RoboDK station: 2026-11-5.rdk

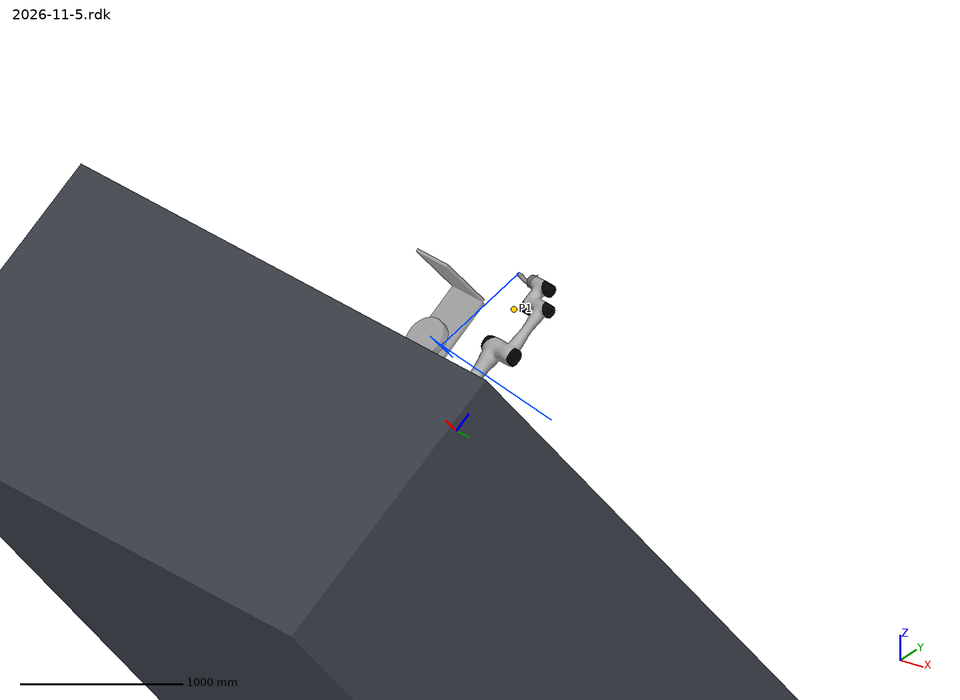
[picture v0: the station drawn from its stored meshes, robots at their saved joint values, targets as dots, program paths as lines]
Station 新建工作站 (1) (saved by RoboDK 5.9.0). Poses are relative to the parent item; angles as X-Y-Z fixed-axis rotations.
Station parameters (name, value as stored): Trace_Render_Style, 0
  - Python program TCP真实运动_升级前备份_20260910_170410 (listed below)
  - Python program 方向角计算 (listed below)
  - Python program test (listed below)
  - Python program 机械臂法兰真实运动_改名修复前_20261014_114144_改名修复前_20261014_114144 (listed below)
  - Python program TCP真实运动_到位复核前备份_20260910_172919 (listed below)
  - Python program TCP真实运动_改名修复前_20261014_114144 (listed below)
  - program _probe_P11 (4 instructions, listed below)
  - Python program 机械臂法兰真实运动 (listed below)
  - Python program TCP仿真 (listed below)
  - Python program TCP真实运动_偏离50版_20261009_142831 (listed below)
  - Python program TCP真实运动_偏离50版_20261009_144043 (listed below)
  - Python program TCP真实运动 (listed below)
  - Python program TCP真实运动_P2P版_修复前_v14w40_20261027 (listed below)
  - Python program TCP真实运动_P2P版_优化前_v14w41_20261027 (listed below)
  - frame Dobot CR5 Base_控制器对齐 at (346.03, 1005.01, 515.52) mm, rotated rx 1.05 ry -48.85 rz -107.35 deg
    - robot Dobot CR5: 6 axes, payload 5 kg, reach 900 mm, repeatability 0.03 mm, weight 23 kg
        modified DH rows (alpha deg, a mm, theta deg, d mm): 0, 0, 0, 147; 90.028, 0.839, 90, 0; -0.44, 427.688, 0, 0; 0.304, 357.005, -90, 140.421; -90.09, 0.126, 0, 115.885; 89.829, 0.736, 180, 104.5
        joint limits [-360, -360, -160, -360, -360, -360] to [360, 360, 160, 360, 360, 360]; home [0, 0, -90, 90, 90, 0]; saved at [0, 0, 0, 0, 0, 0]
      - tool CR5_TCP_126mm, TCP at (0, 0, 126) mm
      - tool _CR5_FLANGE_DIRECT_TEMP, TCP at (0, 0, 0) mm
      - tool _, TCP at (0, 0, 130) mm
      - tool CR5_TCP_130mm, TCP at (0, 0, 130) mm
      - tool _offline_TCP130_test, TCP at (0, 0, 130) mm
      - object  at (0, 0, 0) mm, size 120.1 x 130 x 24.6 mm, geometry from handle130.stl
    - target P1 (joint target) at (-20.1, -241.48, 846.75) mm, rotated rx -90 ry 1.35 rz 179.96 deg; joints [0, -37.451, 84.112, -46.661, 0, 0] of Dobot CR5
    - object  at (0, 0, 0) mm, rotated rx 0 ry -1.35 rz -0.05 deg, size 650 x 650 x 80 mm
    - object  at (0, 0, 0) mm, rotated rx 0 ry -1.35 rz -0.05 deg, size 4000 x 4000 x 2000 mm
    - object  at (0, 223.9, 120) mm, size 450 x 300 x 750 mm, geometry from baffle_semiopen_3face_y300.stl
    - object  at (0, -692.1, 420) mm, rotated rx 90 ry 0 rz 90 deg, size 280 x 280 x 50 mm, geometry from cylinder_R140_H50.stl
  - Python program TCP真实运动_P2P版_16稳定版_替换前_20261104_095940 (listed below)
  - program _TCP仿真_路径预检 (0 instructions, listed below)
  - Python program TCP真实运动_P2P版 (listed below)
  - program 轨迹17_仿真27点 (30 instructions, listed below)
  - object  at (0, 0, 0) mm
  - Python program CR5_零位到P1_上传 (listed below)
  - Python program CR5_首段MoveL_上传 (listed below)
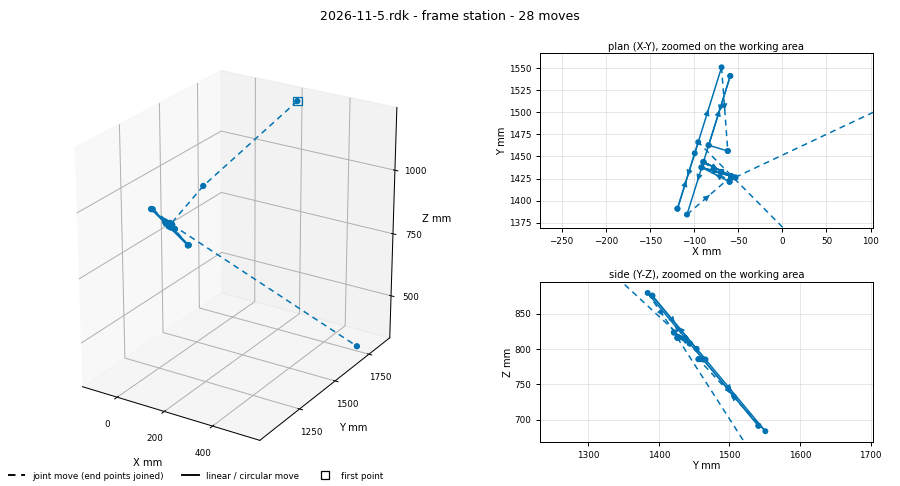
[picture p0: tool path of 2026-11-5.rdk in frame station, 28 of 30 moves have a stored position in this frame; points joined in program order, loops and branches not executed]

--- Python program TCP真实运动_升级前备份_20260910_170410 ---
# -*- coding: utf-8 -*-
"""
RoboDK 实机运动控制（基于 robodk_movej_diag.py 的成功模式）
- 单点：TCP 输入 -> IK 检测 -> MoveL/MoveJ 执行
- 连续轨迹：坐标列表 -> 逐点 IK 检测 -> MoveJ+MoveL 序列
模式：RUNMODE_RUN_ROBOT + robot.Connect()
"""

from robodk.robolink import *
from robodk.robomath import *
import tkinter as tk
from tkinter import ttk, scrolledtext, filedialog
import time
import math
import json

ROBOT_SPEED = 20.0
NL = chr(10)

RDK = Robolink()

def fanuc_to_pose(x, y, z, rx, ry, rz):
    return Fanuc_2_Pose([x, y, z, rx, ry, rz])

def pose_to_fanuc(pose):
    return Pose_2_Fanuc(pose)

# ---- 获取机器人 ----
robot = RDK.Item('', ITEM_TYPE_ROBOT)
if not robot.Valid():
    raise Exception("未找到机器人")

# ---- 全局变量 ----
text_points = None
text_log = None
record_text = None
entries_single = None
entries_joint = None
move_type = None
trajectory_records = []
_connected = False

# ============================================================
# 日志
# ============================================================
def log(s):
    print(s)
    if text_log:
        text_log.insert(tk.END, str(s) + NL)
        text_log.see(tk.END)
        root.update_idletasks()

# ============================================================
# 连接（只连一次，复用）
# ============================================================
def ensure_connected():
    global _connected
    if _connected:
        return True
    try:
        robot.Connect()
        time.sleep(1.5)
        status, msg = robot.ConnectedState()
        log("连接状态: %s, %s" % (status, msg))
        RDK.setRunMode(RUNMODE_RUN_ROBOT)
        log("RunMode: %s" % RDK.RunMode())
        if status < 0:
            _connected = False
            log("机器人连接未建立，状态=%s：%s" % (status, msg))
            return False
        _connected = True
        return True
    except Exception as e:
        log("连接失败: %s" % e)
        return False

# ============================================================
# 解析坐标
# ============================================================
def parse_points():
    if not text_points:
        return []
    raw = text_points.get("1.0", tk.END)
    points = []
    for line in raw.strip().split(NL):
        line = line.strip()
        if not line or line.startswith("#"):
            continue
        try:
            vals = [float(v.strip()) for v in line.split(",")]
            if len(vals) >= 6:
                points.append(vals[:6])
        except ValueError:
            pass
    return points

# ============================================================
# 读取当前位置
# ============================================================
def read_current(entries=None):
    try:
        pose = robot.Pose()
        v = pose_to_fanuc(pose)
        log("")
        log("当前 TCP：X=%.3f Y=%.3f Z=%.3f Rx=%.3f Ry=%.3f Rz=%.3f" % tuple(v[:6]))
    except Exception as e:
        log("读取失败：%s" % e)

def fill_current(entries=None):
    try:
        pose = robot.Pose()
        v = pose_to_fanuc(pose)
        if entries:
            for e, val in zip(entries, v):
                e.delete(0, tk.END)
                e.insert(0, "%.3f" % val)
        log("当前 TCP 已填入")
    except Exception as e:
        log("读取失败：%s" % e)

# ============================================================
# IK 检测
# 注意：SolveIK 显式使用当前 Tool + Reference，和 MoveL/MoveJ 保持一致。
# ============================================================
def check_ik_single(entries=None):
    if not entries:
        return
    try:
        values = [float(e.get()) for e in entries]
    except ValueError:
        log("输入无效")
        return

    x, y, z, rx, ry, rz = values
    target = fanuc_to_pose(x, y, z, rx, ry, rz)
    log("")
    log("目标：X=%.3f Y=%.3f Z=%.3f Rx=%.3f Ry=%.3f Rz=%.3f" % (x, y, z, rx, ry, rz))

    try:
        tool_pose = robot.PoseTool()
        frame_pose = robot.PoseFrame()
        joints = robot.SolveIK(target, tool=tool_pose, reference=frame_pose)
        if joints is None:
            log("IK 不可达")
        else:
            q = joints.list()
            if len(q) < 6:
                log("IK 返回关节数量异常：%d，原始数据=%r" % (len(q), q))
                return
            log("IK 可达")
            log("  关节：J1=%.2f J2=%.2f J3=%.2f J4=%.2f J5=%.2f J6=%.2f" % tuple(q[:6]))
    except Exception as e:
        log("检测失败：%s" % e)

def check_all_ik():
    points = parse_points()
    if not points:
        log("没有有效点")
        return

    log("")
    log("========== 检测全部 %d 个点 ==========" % len(points))
    all_ok = True
    for i, p in enumerate(points):
        try:
            target = fanuc_to_pose(*p)
            joints = robot.SolveIK(target, tool=robot.PoseTool(), reference=robot.PoseFrame())
            if joints is None:
                log("  P%d: 不可达" % (i+1))
                all_ok = False
            else:
                q = joints.list()
                if len(q) < 6:
                    raise ValueError("IK 返回关节数量异常: %d, raw=%r" % (len(q), q))
                log("  P%d: 可达  J1=%.1f J2=%.1f J3=%.1f J4=%.1f J5=%.1f J6=%.1f" % (i+1, *q[:6]))
        except Exception as e:
            log("  P%d: 检测失败 %s" % (i+1, e))
            all_ok = False
    if all_ok:
        log("全部 %d 个点可达" % len(points))
    else:
        log("存在不可达点，执行时会跳过")

# ============================================================
# 执行单点
# ============================================================
def execute_single(entries=None, mtype="MoveL"):
    if not entries:
        return
    try:
        values = [float(e.get()) for e in entries]
    except ValueError:
        log("输入无效")
        return

    x, y, z, rx, ry, rz = values
    target = fanuc_to_pose(x, y, z, rx, ry, rz)
    log("")
    log("目标：X=%.3f Y=%.3f Z=%.3f Rx=%.3f Ry=%.3f Rz=%.3f" % (x, y, z, rx, ry, rz))

    try:
        tool_pose = robot.PoseTool()
        frame_pose = robot.PoseFrame()
        joints = robot.SolveIK(target, tool=tool_pose, reference=frame_pose)
        if joints is None:
            log("IK 不可达，取消执行")
            return
        q = joints.list()
        if len(q) < 6:
            log("IK 返回关节数量异常：%d，取消执行；原始数据=%r" % (len(q), q))
            return
        log("IK 可达：J1=%.2f J2=%.2f J3=%.2f J4=%.2f J5=%.2f J6=%.2f" % tuple(q[:6]))
    except Exception as e:
        log("IK 检查失败：%s" % e)
        return

    if not ensure_connected():
        return

    try:
        robot.setPoseFrame(robot.PoseFrame())
        robot.setPoseTool(robot.PoseTool())
        robot.setSpeed(ROBOT_SPEED)
        log("发送 %s..." % mtype)
        if mtype == "MoveJ":
            robot.MoveJ(target)
        else:
            robot.MoveL(target)
        log("执行完成")
    except Exception as e:
        log("失败: %s: %s" % (type(e).__name__, e))

# ============================================================
# 连续运动：选项卡3直接输入 TCP / 关节点，逐点检查后加入轨迹
# ============================================================
trajectory_records = []
record_text = None
traj_entries = None
traj_type = None
singular_var = None
j6_direction_var = None


def _parse_six_from_entries(entries, label):
    if not entries or len(entries) != 6:
        log("%s输入框异常：需要 6 个值" % label)
        return None
    try:
        vals = [float(e.get().strip()) for e in entries]
    except (ValueError, AttributeError):
        log("%s输入无效：6 个值必须全部为数字" % label)
        return None
    if not all(math.isfinite(v) for v in vals):
        log("%s输入无效：不能包含 NaN 或无穷值" % label)
        return None
    return vals


def _check_tcp_reachable(vals):
    """检查单个 TCP 点 IK 是否可达，返回 (True, target, joints)。"""
    try:
        target = fanuc_to_pose(*vals)
        tool_pose = robot.PoseTool()
        frame_pose = robot.PoseFrame()
        joints = robot.SolveIK(target, tool=tool_pose, reference=frame_pose)

        if joints is None:
            log("TCP IK：不可达")
            return False, None, None

        q = joints.list()
        if len(q) < 6:
            log("TCP IK：返回关节数量异常：%r" % q)
            return False, None, None

        log("TCP IK：可达")
        log("  IK关节：J1=%.2f J2=%.2f J3=%.2f J4=%.2f J5=%.2f J6=%.2f" % tuple(q[:6]))
        return True, target, q[:6]
    except Exception as e:
        log("TCP IK 检查失败：%s: %s" % (type(e).__name__, e))
        return False, None, None


def _check_tcp_segment_continuous(prev_vals, curr_vals, segment_index, samples=20):
    """检查前一个 TCP 点到当前 TCP 点之间的整段插补路径 IK 连续可达性。

    暂不考虑障碍物，只对 TCP 位姿做线性插值，并对每个采样位姿执行 SolveIK。
    起点和终点也包含在采样检查中。
    """
    if prev_vals is None:
        return True

    log("开始检查 P%d -> P%d 的 TCP 连续 IK（%d 个采样点）" %
        (segment_index - 1, segment_index, samples + 1))

    tool_pose = robot.PoseTool()
    frame_pose = robot.PoseFrame()

    for k in range(samples + 1):
        t = float(k) / float(samples)
        vals = [prev_vals[i] + (curr_vals[i] - prev_vals[i]) * t for i in range(6)]
        try:
            pose = fanuc_to_pose(*vals)
            joints = robot.SolveIK(pose, tool=tool_pose, reference=frame_pose)
            if joints is None:
                log("  P%d -> P%d：第 %d/%d 个采样点 IK 不可达，t=%.3f" %
                    (segment_index - 1, segment_index, k + 1, samples + 1, t))
                log("  TCP：X=%.3f Y=%.3f Z=%.3f Rx=%.3f Ry=%.3f Rz=%.3f" % tuple(vals))
                return False
            q = joints.list()
            if len(q) < 6:
                log("  P%d -> P%d：第 %d 个采样点 IK 返回异常：%r" %
                    (segment_index - 1, segment_index, k + 1, q))
                return False
        except Exception as e:
            log("  P%d -> P%d：第 %d 个采样点 IK 检查失败：%s: %s" %
                (segment_index - 1, segment_index, k + 1, type(e).__name__, e))
            return False

    log("P%d -> P%d：连续 IK 检查通过" % (segment_index - 1, segment_index))
    return True


def _check_joint_reachable(q):
    """兼容旧代码：关节点不做可达性/限位检查，输入合法即可加入。"""
    return True


def refresh_record_list():
    if record_text is None:
        return

    record_text.delete("1.0", tk.END)

    for i, rec in enumerate(trajectory_records, 1):
        kind = rec["type"]
        vals = rec["values"]

        if kind == "TCP":
            mark = " [J6特异点 %s180°]" % ("+" if rec.get("j6_delta", 180) >= 0 else "-") if rec.get("singular", False) else ""
            record_text.insert(
                tk.END,
                "P%-3d [TCP]%s   X=%9.3f Y=%9.3f Z=%9.3f Rx=%8.3f Ry=%8.3f Rz=%8.3f%s" %
                (i, mark, *vals, NL)
            )
        else:
            record_text.insert(
                tk.END,
                "P%-3d [JNT]   J1=%8.3f J2=%8.3f J3=%8.3f J4=%8.3f J5=%8.3f J6=%8.3f%s" %
                (i, *vals, NL)
            )


def add_and_check_trajectory_point():
    """
    选项卡3逐点输入：
    - 普通 TCP：立即做端点 IK，并检查与前一个普通 TCP 点之间的连续 IK。
    - TCP 末端特异点：跳过 IK；要求与前一个普通 TCP 点 XYZ 相同，执行时仅 J6 转 ±180°。
    - 关节：不做 IK/限位检查，只将角度规范到 (-180°, 180°]。
    注意：这些检查只在“加入点”时完成；正式实机执行时不再做轨迹预检。
    """
    kind = traj_type.get()
    vals = _parse_six_from_entries(traj_entries, kind)
    if vals is None:
        return

    log("")
    log("========== 检查连续运动第 %d 点 ==========" % (len(trajectory_records) + 1))

    is_singular = bool(singular_var.get()) if (kind == "TCP" and singular_var is not None) else False
    j6_delta = int(j6_direction_var.get()) if (j6_direction_var is not None) else 180

    if kind == "TCP" and is_singular:
        if not trajectory_records:
            log("末端特异点不能作为第一个点：需要先有一个起始运动点。")
            return
        prev = trajectory_records[-1]
        if prev["type"] != "TCP" or prev.get("singular", False):
            log("末端特异点前一项必须是普通 TCP 点。")
            return
        prev_vals = prev["values"]
        pos_err = math.sqrt(sum((vals[k] - prev_vals[k]) ** 2 for k in range(3)))
        if pos_err > 1e-3:
            log("末端特异点未加入：XYZ 必须与前一个普通 TCP 点相同。")
            log("  与前一点位置差：%.6f mm" % pos_err)
            return
        try:
            target = fanuc_to_pose(*vals)
        except Exception as e:
            log("末端特异点姿态转换失败：%s: %s" % (type(e).__name__, e))
            return

        trajectory_records.append({
            "type": "TCP", "values": vals[:], "target": target, "joints": None,
            "singular": True, "j6_delta": j6_delta,
        })
        log("P%d [TCP-特异点]：已加入，跳过 IK。" % len(trajectory_records))
        log("  执行时保持 J1~J5 不变，仅让 J6 转 %+d°。" % j6_delta)
        if singular_var is not None:
            singular_var.set(False)
        refresh_record_list()
        return

    if kind == "TCP":
        ok, target, joints = _check_tcp_reachable(vals)
        if not ok:
            log("该 TCP 点未加入轨迹。")
            return

        # 只在点加入阶段检查连续 IK；实机正式执行时不再重复预检。
        if trajectory_records and trajectory_records[-1]["type"] == "TCP" and not trajectory_records[-1].get("singular", False):
            prev_vals = trajectory_records[-1]["values"]
            segment_no = len(trajectory_records) + 1
            if not _check_tcp_segment_continuous(prev_vals, vals, segment_no, samples=20):
                log("P%d [TCP]：上一普通 TCP 点到当前点的连续 IK 检查失败，该点未加入轨迹。" % segment_no)
                return

        trajectory_records.append({
            "type": "TCP", "values": vals[:], "target": target, "joints": joints,
            "singular": False, "j6_delta": 0,
        })
        log("P%d [TCP]：检查通过，已加入连续运动。" % len(trajectory_records))
    else:
        corrected = []
        for v in vals:
            v = ((v + 180.0) % 360.0) - 180.0
            if v <= -180.0:
                v = 180.0
            corrected.append(v)
        if corrected != vals:
            log("关节点角度已自动纠正到 (-180°, 180°]：")
            log("  原始：" + "  ".join("J%d=%+.3f°" % (i + 1, vals[i]) for i in range(6)))
            log("  修正：" + "  ".join("J%d=%+.3f°" % (i + 1, corrected[i]) for i in range(6)))
        trajectory_records.append({
            "type": "JOINT", "values": corrected[:], "target": None, "joints": corrected[:],
            "singular": False, "j6_delta": 0,
        })
        log("P%d [JNT]：未做 IK 检查，角度规范化后已加入连续运动。" % len(trajectory_records))

    refresh_record_list()


def _write_values_to_traj_entries(values, label):
    if not traj_entries or len(traj_entries) != 6:
        log("连续运动输入框异常：无法写入当前%s" % label)
        return False
    for e, val in zip(traj_entries, values[:6]):
        e.delete(0, tk.END)
        e.insert(0, "%.3f" % float(val))
    log("当前%s已写入选项卡3输入框" % label)
    return True


def read_current_tcp_to_traj():
    """读取当前 RoboDK TCP，并写入选项卡3的 TCP 输入框。"""
    try:
        pose = robot.Pose()
        vals = pose_to_fanuc(pose)
        log("========== 读取当前 TCP -> 选项卡3 ==========")
        log("X=%+.3f Y=%+.3f Z=%+.3f Rx=%+.3f Ry=%+.3f Rz=%+.3f" % tuple(vals))
        if traj_type.get() != "TCP":
            traj_type.set("TCP")
            _update_traj_labels_and_defaults()
        return _write_values_to_traj_entries(vals, "TCP")
    except Exception as e:
        log("读取当前 TCP 失败：%s: %s" % (type(e).__name__, e))
        return False


def read_current_joints_to_traj():
    """读取 RoboDK Robot Item 当前关节，并写入选项卡3的关节输入框。"""
    q = read_current_joints(None)
    if q is None or len(q) < 6:
        return False
    log("========== 读取当前关节 -> 选项卡3 ==========")
    if traj_type.get() != "JOINT":
        traj_type.set("JOINT")
        _update_traj_labels_and_defaults()
    return _write_values_to_traj_entries(q, "关节")


def clear_trajectory_input():
    if not traj_entries:
        return

    for e in traj_entries:
        e.delete(0, tk.END)

    if traj_type.get() == "TCP":
        defaults = ["0.000", "-241.500", "1047.000", "-90.000", "0.000", "180.000"]
    else:
        defaults = ["0.000"] * 6

    for e, val in zip(traj_entries, defaults):
        e.insert(0, val)




def import_trajectory():
    """
    从仿真程序导出的 JSON 轨迹文件导入到实机连续运动列表。

    重要：这里不做连续轨迹预检，不做 MoveJ TCP 轨迹预检。
    普通 TCP 如果 JSON 中没有保存 IK 关节，则只针对该点单独 SolveIK，
    用于得到实机执行所需的目标关节；这不是连续轨迹预检。
    """
    filepath = filedialog.askopenfilename(
        title="导入仿真轨迹",
        defaultextension=".json",
        filetypes=[("JSON 轨迹文件", "*.json"), ("所有文件", "*.*")]
    )
    if not filepath:
        return

    try:
        with open(filepath, "r", encoding="utf-8") as f:
            data = json.load(f)

        if not isinstance(data, list):
            raise ValueError("轨迹文件顶层必须是列表。")

        imported = []
        for idx, item in enumerate(data, 1):
            if not isinstance(item, dict):
                raise ValueError("P%d 不是对象格式。" % idx)

            kind = str(item.get("type", "")).upper()
            if kind == "JNT":
                kind = "JOINT"
            if kind not in ("TCP", "JOINT"):
                raise ValueError("P%d type 不支持：%r" % (idx, item.get("type")))

            values = item.get("values")
            if not isinstance(values, list) or len(values) != 6:
                raise ValueError("P%d values 必须是长度为6的列表。" % idx)
            try:
                values = [float(v) for v in values]
            except (TypeError, ValueError):
                raise ValueError("P%d values 必须全部为数字。" % idx)
            if not all(math.isfinite(v) for v in values):
                raise ValueError("P%d values 不能包含 NaN 或无穷值。" % idx)

            is_singular = bool(item.get("singular", False)) and kind == "TCP"
            j6_delta = int(item.get("j6_delta", 180)) if is_singular else 0
            if is_singular and j6_delta not in (-180, 180):
                raise ValueError("P%d 特异点 j6_delta 只能是 +180 或 -180。" % idx)

            if kind == "JOINT":
                # 与手动输入保持一致：自动规范到 (-180,180]。
                corrected = []
                for v in values:
                    v = ((v + 180.0) % 360.0) - 180.0
                    if v <= -180.0:
                        v = 180.0
                    corrected.append(v)
                values = corrected
                imported.append({
                    "type": "JOINT", "values": values, "target": None,
                    "joints": values[:], "singular": False, "j6_delta": 0
                })
                continue

            target = fanuc_to_pose(*values)

            if is_singular:
                # 特异点严格要求前一项为普通 TCP，且 XYZ 相同。
                if not imported:
                    raise ValueError("P%d 末端特异点不能作为第一个点。" % idx)
                prev = imported[-1]
                if prev["type"] != "TCP" or prev.get("singular", False):
                    raise ValueError("P%d 末端特异点前一项必须是普通 TCP。" % idx)
                pos_err = math.sqrt(sum((values[k] - prev["values"][k]) ** 2 for k in range(3)))
                if pos_err > 1e-3:
                    raise ValueError("P%d 末端特异点 XYZ 必须与前一个普通 TCP 相同，位置差 %.6f mm。" % (idx, pos_err))
                imported.append({
                    "type": "TCP", "values": values[:], "target": target,
                    "joints": None, "singular": True, "j6_delta": j6_delta
                })
                continue

            # 优先使用文件中可能保存的 IK；当前仿真脚本的 JSON 通常没有 joints，
            # 因此回退到“单点 SolveIK”，仅为了得到实机 MoveJ/MoveL 所需目标关节。
            q = item.get("joints")
            if isinstance(q, list) and len(q) >= 6:
                try:
                    q = [float(v) for v in q[:6]]
                    if not all(math.isfinite(v) for v in q):
                        q = None
                except (TypeError, ValueError):
                    q = None

            if q is None:
                joints = robot.SolveIK(
                    target, tool=robot.PoseTool(), reference=robot.PoseFrame()
                )
                if joints is None:
                    raise ValueError("P%d 普通 TCP 单点 IK 无解，无法导入。" % idx)
                q = joints.list()
                if q is None or len(q) < 6:
                    raise ValueError("P%d 普通 TCP IK 返回关节数量异常：%r" % (idx, q))
                q = [float(v) for v in q[:6]]

            imported.append({
                "type": "TCP", "values": values[:], "target": target,
                "joints": q[:], "singular": False, "j6_delta": 0
            })

        trajectory_records.clear()
        trajectory_records.extend(imported)
        refresh_record_list()
        log("")
        log("========== 导入仿真轨迹 ==========")
        log("文件：%s" % filepath)
        log("已导入 %d 个轨迹点。" % len(imported))
        log("连续轨迹预检：未执行（按实机程序设计）。")
        log("普通 TCP：仅在缺少保存IK时进行单点 SolveIK；不进行连续段预检。")
        log("末端特异点：跳过IK，仅保留 J6 ±180° 标记。")
        log("================================")
    except Exception as e:
        log("轨迹导入失败：%s: %s" % (type(e).__name__, e))

def delete_last_record():
    if trajectory_records:
        rec = trajectory_records.pop()
        refresh_record_list()
        log("已删除最后一点：P%d [%s]" %
            (len(trajectory_records) + 1, rec["type"]))
    else:
        log("当前没有可删除的连续运动点")


def clear_records():
    trajectory_records.clear()
    refresh_record_list()
    log("连续运动点列表已清空")


def execute_recorded_trajectory():
    """
    实机执行选项卡3轨迹。

    重要：不做仿真轨迹预检。TCP 的 IK/连续 IK 已在“检查并加入当前点”阶段完成，
    实机这里只负责按仿真已经验证过的顺序执行。

    普通 TCP：第一个 TCP MoveJ，后续普通 TCP 优先 MoveL；MoveL 失败后直接用已经保存的 IK 关节 MoveJ 兜底。
    末端特异点：跳过 IK，读取当前 RoboDK Robot Item 关节，仅 J6 转 ±180°。
    特异点后的普通 TCP：重新使用该普通 TCP 自己保存的 IK，正常 MoveL。
    关节点：直接 MoveJ。
    StoppedError: Robot not connected：继续视为本段结束标志。
    """
    if not trajectory_records:
        log("没有已检查通过的运动点，请先在选项卡3输入并加入点。")
        return

    log("")
    log("========== 执行实机连续运动：%d 个点 ==========" % len(trajectory_records))
    log("轨迹预检：跳过（已在仿真/加入点阶段完成）")

    if not ensure_connected():
        log("连续运动取消：机器人未连接")
        return

    try:
        RDK.setRunMode(RUNMODE_RUN_ROBOT)
        robot.setPoseFrame(robot.PoseFrame())
        robot.setPoseTool(robot.PoseTool())
        robot.setSpeed(ROBOT_SPEED)

        tcp_count = 0
        completed_count = 0

        for i, rec in enumerate(trajectory_records, 1):
            kind = rec["type"]
            vals = rec["values"]
            is_singular = bool(rec.get("singular", False))
            j6_delta = int(rec.get("j6_delta", 180))

            if kind == "TCP" and is_singular:
                move_name = "J6特异点"
            elif kind == "TCP":
                move_name = "MoveJ" if tcp_count == 0 else "MoveL"
            else:
                move_name = "MoveJ"

            log("")
            log("---- 开始执行 P%d [%s] -> %s ----" % (i, kind, move_name))

            try:
                if kind == "TCP":
                    if is_singular:
                        # 特异点：当前 RoboDK Robot Item 关节作为起点，保持 J1~J5，仅改变 J6。
                        current_q = list(robot.SimulatorJoints())
                        if len(current_q) < 6:
                            raise RuntimeError("特异点：RoboDK SimulatorJoints 返回关节数量不足6个：%r" % current_q)
                        current_q = current_q[:6]
                        q_special = current_q[:]
                        q_special[5] += float(j6_delta)
                        # 保持与前面关节点规范一致，避免无意义多圈累加。
                        q_special[5] = ((q_special[5] + 180.0) % 360.0) - 180.0
                        if q_special[5] <= -180.0:
                            q_special[5] = 180.0
                        log("P%d [TCP-特异点]：J6 %.3f° -> %.3f°，J1~J5保持不变" %
                            (i, current_q[5], q_special[5]))
                        robot.MoveJ(q_special)
                        tcp_count += 1
                    elif tcp_count == 0:
                        # 首个普通TCP：使用加入阶段已经得到的IK关节，避免再次SolveIK。
                        q = rec.get("joints")
                        if q is None or len(q) < 6:
                            raise RuntimeError("P%d：缺少已保存的 TCP IK 关节解。" % i)
                        robot.MoveJ(q[:6])
                        tcp_count += 1
                    else:
                        # 后续普通TCP：优先 MoveL。
                        target = rec.get("target")
                        q = rec.get("joints")
                        if target is None or q is None or len(q) < 6:
                            raise RuntimeError("P%d：缺少已保存的 TCP 目标位姿或 IK 关节解。" % i)
                        try:
                            robot.MoveL(target)
                        except Exception as e_l:
                            # 仿真已经检查过 MoveJ 的 TCP 轨迹，因此实机不再重复预检，直接用已验证的 IK 解兜底。
                            log("P%d [TCP] -> MoveL 失败：%s: %s" % (i, type(e_l).__name__, e_l))
                            log("P%d [TCP] -> 直接使用仿真已验证的 IK 关节解执行 MoveJ 兜底。" % i)
                            robot.MoveJ(q[:6])

                else:
                    q = rec["values"][:6]
                    robot.MoveJ(q)

                completed_count += 1
                log("P%d [%s] -> %s 返回正常，进入下一段。" % (i, kind, move_name))

            except Exception as e:
                err_type = type(e).__name__
                err_text = str(e)
                if err_type == "StoppedError" and "Robot not connected" in err_text:
                    completed_count += 1
                    log("P%d [%s] -> %s 已结束。" % (i, kind, move_name))
                    log("收到结束标志：StoppedError: Robot not connected")
                    log("将该报错视为本段运动结束，继续执行下一段。")
                    continue

                log("P%d [%s] -> %s 执行失败：%s: %s" %
                    (i, kind, move_name, err_type, err_text))
                log("非预期错误，停止后续连续运动。")
                return

        log("")
        log("========== 实机连续运动执行完成：%d/%d 段 ==========" %
            (completed_count, len(trajectory_records)))

    except Exception as e:
        log("连续运动初始化失败：%s: %s" % (type(e).__name__, e))


# 保留旧函数名，避免其他代码调用失效。
def execute_trajectory():
    execute_recorded_trajectory()


# ============================================================
# 实机关节运动
# ============================================================
def _joint_values_from_entries(entries):
    """从 GUI 读取 J1~J6 目标角度。单位：deg。"""
    if not entries or len(entries) != 6:
        log("目标关节输入框异常：需要 J1~J6 共 6 个")
        return None
    try:
        q = [float(e.get().strip()) for e in entries]
    except (ValueError, AttributeError):
        log("目标关节输入无效：J1~J6 必须全部填写数字")
        return None
    if not all(math.isfinite(v) for v in q):
        log("目标关节输入无效：不能包含 NaN 或无穷值")
        return None
    return q


def read_current_joints(entries=None):
    """读取 RoboDK Robot Item 当前关节值，并可直接填入 J1~J6 输入框。
    注意：这里读取的是 RoboDK 当前 Robot Item 的关节状态，不调用 CR5 控制器 GetAngle。
    """
    try:
        joints = robot.SimulatorJoints()
        q = list(joints) if hasattr(joints, "__iter__") else [joints]
        if len(q) < 6:
            log("读取当前关节失败：SimulatorJoints 返回 %r" % (q,))
            log("请确认 RoboDK 窗口中的机器人已经连接并显示实时关节角度。")
            return None

        q = q[:6]
        log("")
        log("========== RoboDK 当前关节 ==========")
        log("J1=%+.3f°  J2=%+.3f°  J3=%+.3f°" % tuple(q[:3]))
        log("J4=%+.3f°  J5=%+.3f°  J6=%+.3f°" % tuple(q[3:]))

        if entries and len(entries) == 6:
            for e, val in zip(entries, q):
                e.delete(0, tk.END)
                e.insert(0, "%.3f" % val)
            log("当前关节已填入 J1~J6 输入框")

        return q
    except Exception as e:
        log("读取 RoboDK 当前关节失败：%s: %s" % (type(e).__name__, e))
        return None


def fill_current_joints(entries=None):
    """当前 RoboDK 关节 -> 目标关节输入框。"""
    return read_current_joints(entries)


def execute_joint_target(entries=None):
    """按 GUI 输入的 J1~J6 目标角度直接执行实机 MoveJ，不经过 TCP/IK。"""
    q = _joint_values_from_entries(entries)
    if q is None:
        return

    log("")
    log("========================================")
    log("====== 实机指定关节角度 MoveJ ======")
    log("目标：J1=%+.3f°  J2=%+.3f°  J3=%+.3f°" % tuple(q[:3]))
    log("      J4=%+.3f°  J5=%+.3f°  J6=%+.3f°" % tuple(q[3:]))
    log("运动速度：%.1f" % ROBOT_SPEED)
    log("控制方式：RoboDK Robot Item -> RUNMODE_RUN_ROBOT -> MoveJ(q)")

    if not ensure_connected():
        log("实机关节运动取消：机器人未连接")
        return

    try:
        RDK.setRunMode(RUNMODE_RUN_ROBOT)
        log("RunMode：%s" % RDK.RunMode())
        robot.setSpeed(ROBOT_SPEED)
        log("发送 MoveJ 目标：%r" % q)
        robot.MoveJ(q)
        log("MoveJ 命令已发送，目标关节角度：%r" % q)
        log("========================================")
    except Exception as e:
        log("实机 MoveJ 失败：%s: %s" % (type(e).__name__, e))


def clear_joint_target(entries=None):
    if not entries:
        return
    for e in entries:
        e.delete(0, tk.END)
        e.insert(0, "0.000")
    log("目标关节输入已清零")

# ============================================================
# GUI
# ============================================================
root = tk.Tk()
root.title("RoboDK - 机械臂运动控制")
root.geometry("1200x750")
root.resizable(True, True)

tk.Label(root, text="Dobot CR5 运动控制", font=("Microsoft YaHei", 16, "bold")).pack(pady=10)

notebook = ttk.Notebook(root)
notebook.pack(fill=tk.BOTH, expand=True, padx=10, pady=5)

# ---- 选项卡 1：单点运动 ----
tab_single = ttk.Frame(notebook)
notebook.add(tab_single, text="单点运动")

frame_coord = tk.LabelFrame(tab_single, text="目标 TCP（Fanuc 格式）")
frame_coord.pack(fill=tk.X, padx=10, pady=10)

names = ["X (mm)", "Y (mm)", "Z (mm)", "Rx (deg)", "Ry (deg)", "Rz (deg)"]
defaults = ["0.000", "-241.500", "1047.000", "-90.000", "0.000", "180.000"]
entries_single = []

for i in range(6):
    tk.Label(frame_coord, text=names[i]).grid(row=0, column=i*2, padx=5, pady=10)
    e = tk.Entry(frame_coord, width=12)
    e.insert(0, defaults[i])
    e.grid(row=0, column=i*2+1, padx=5, pady=10)
    entries_single.append(e)

frame_mtype = tk.Frame(tab_single)
frame_mtype.pack(fill=tk.X, padx=10, pady=5)
move_type = tk.StringVar(value="MoveL")
tk.Radiobutton(frame_mtype, text="MoveL (直线)", variable=move_type, value="MoveL").pack(side=tk.LEFT, padx=10)
tk.Radiobutton(frame_mtype, text="MoveJ (关节)", variable=move_type, value="MoveJ").pack(side=tk.LEFT, padx=10)

btn_single_frame = tk.Frame(tab_single)
btn_single_frame.pack(fill=tk.X, padx=10, pady=5)

def _read_current():
    read_current(entries_single)
def _fill_current():
    fill_current(entries_single)
def _check_ik():
    check_ik_single(entries_single)
def _exec_single():
    execute_single(entries_single, move_type.get())

tk.Button(btn_single_frame, text="读取当前 TCP", command=_read_current, width=15).pack(side=tk.LEFT, padx=3)
tk.Button(btn_single_frame, text="当前 TCP -> 输入框", command=_fill_current, width=20).pack(side=tk.LEFT, padx=3)
tk.Button(btn_single_frame, text="检测可达性", command=_check_ik, width=15, bg="#2196F3", fg="white").pack(side=tk.LEFT, padx=3)
tk.Button(btn_single_frame, text="执行运动", command=_exec_single, width=20,
          font=("Microsoft YaHei", 10, "bold"), bg="#4CAF50", fg="white").pack(side=tk.LEFT, padx=3)


# ---- 选项卡 2：目标关节运动（实机） ----
tab_joint = ttk.Frame(notebook)
notebook.add(tab_joint, text="目标关节运动")

frame_joint = tk.LabelFrame(tab_joint, text="目标关节（deg）")
frame_joint.pack(fill=tk.X, padx=10, pady=10)

joint_names = ["J1 (deg)", "J2 (deg)", "J3 (deg)", "J4 (deg)", "J5 (deg)", "J6 (deg)"]
joint_defaults = ["0.000", "0.000", "0.000", "0.000", "0.000", "0.000"]
entries_joint = []

for i in range(6):
    tk.Label(frame_joint, text=joint_names[i]).grid(row=0, column=i*2, padx=5, pady=10)
    e = tk.Entry(frame_joint, width=12)
    e.insert(0, joint_defaults[i])
    e.grid(row=0, column=i*2+1, padx=5, pady=10)
    entries_joint.append(e)

btn_joint_frame = tk.Frame(tab_joint)
btn_joint_frame.pack(fill=tk.X, padx=10, pady=8)

def _read_current_joint_values():
    read_current_joints(entries_joint)

def _fill_current_joints():
    fill_current_joints(entries_joint)

def _exec_joint():
    execute_joint_target(entries_joint)

def _zero_joints():
    clear_joint_target(entries_joint)

tk.Button(btn_joint_frame, text="读取当前关节", command=_read_current_joint_values, width=14).pack(side=tk.LEFT, padx=3)
tk.Button(btn_joint_frame, text="当前关节 -> 输入框", command=_fill_current_joints, width=20).pack(side=tk.LEFT, padx=3)
tk.Button(btn_joint_frame, text="执行指定关节 MoveJ", command=_exec_joint, width=24,
          font=("Microsoft YaHei", 10, "bold"), bg="#FF9800", fg="white").pack(side=tk.LEFT, padx=3)
tk.Button(btn_joint_frame, text="清零", command=_zero_joints, width=10).pack(side=tk.LEFT, padx=3)

tk.Label(tab_joint,
         text="输入 J1~J6 目标角度（deg），点击“执行指定关节 MoveJ”直接控制实机；不经过 TCP、Fanuc 转换或 IK。",
         fg="#555555").pack(anchor=tk.W, padx=15, pady=5)
tk.Label(tab_joint,
         text="安全提示：首次测试建议只改变一个关节、改变 5~10°，确认方向和角度定义正确后再进行大角度运动。",
         fg="#C62828").pack(anchor=tk.W, padx=15, pady=2)

# ---- 选项卡 3：连续运动 ----
tab_traj = ttk.Frame(notebook)
notebook.add(tab_traj, text="连续运动")

frame_traj_input = tk.LabelFrame(
    tab_traj,
    text="连续运动点输入：每次输入 1 个 TCP 点或 1 组关节角度，点击“检查并加入”"
)
frame_traj_input.pack(fill=tk.X, padx=10, pady=10)

type_frame = tk.Frame(frame_traj_input)
type_frame.pack(fill=tk.X, padx=8, pady=5)

tk.Label(type_frame, text="点类型：").pack(side=tk.LEFT, padx=3)

traj_type = tk.StringVar(value="TCP")
tk.Radiobutton(
    type_frame, text="TCP（X,Y,Z,Rx,Ry,Rz）",
    variable=traj_type, value="TCP"
).pack(side=tk.LEFT, padx=8)

tk.Radiobutton(
    type_frame, text="关节（J1~J6）",
    variable=traj_type, value="JOINT"
).pack(side=tk.LEFT, padx=8)

traj_names_tcp = ["X", "Y", "Z", "Rx", "Ry", "Rz"]
traj_names_joint = ["J1", "J2", "J3", "J4", "J5", "J6"]

traj_entries = []

# ---- 末端特异点设置 ----
singular_var = tk.BooleanVar(value=False)
j6_direction_var = tk.IntVar(value=180)

singular_frame = tk.Frame(frame_traj_input)
singular_frame.pack(fill=tk.X, padx=8, pady=3)

tk.Checkbutton(
    singular_frame,
    text="末端特异点（跳过IK，仅J6转180°）",
    variable=singular_var
).pack(side=tk.LEFT, padx=3)

tk.Label(singular_frame, text="J6方向：").pack(side=tk.LEFT, padx=(15, 3))
tk.Radiobutton(singular_frame, text="+180°", variable=j6_direction_var, value=180).pack(side=tk.LEFT, padx=3)
tk.Radiobutton(singular_frame, text="-180°", variable=j6_direction_var, value=-180).pack(side=tk.LEFT, padx=3)

# 输入框单独放在 grid 子容器中。
# frame_traj_input 本身使用 pack 管理子控件，不能再直接对它的子控件使用 grid。
traj_value_frame = tk.Frame(frame_traj_input)
traj_value_frame.pack(fill=tk.X, padx=8, pady=5)

for i in range(6):
    tk.Label(
        traj_value_frame,
        text=traj_names_tcp[i]
    ).grid(row=0, column=i * 2, padx=3, pady=8)

    e = tk.Entry(traj_value_frame, width=12)
    e.grid(row=0, column=i * 2 + 1, padx=4, pady=8)
    traj_entries.append(e)

# 默认先按 TCP 输入显示
tcp_defaults = ["0.000", "-241.500", "1047.000", "-90.000", "0.000", "180.000"]
for e, val in zip(traj_entries, tcp_defaults):
    e.insert(0, val)


def _update_traj_labels_and_defaults():
    """切换 TCP/关节输入时，更新标签和默认值。"""
    names = traj_names_tcp if traj_type.get() == "TCP" else traj_names_joint
    defaults = (
        tcp_defaults
        if traj_type.get() == "TCP"
        else ["0.000"] * 6
    )

    for i, e in enumerate(traj_entries):
        # grid 上的 Label 位于当前列
        for widget in traj_value_frame.grid_slaves(row=0, column=i * 2):
            widget.configure(text=names[i])

        e.delete(0, tk.END)
        e.insert(0, defaults[i])


tk.Radiobutton(
    type_frame, text="TCP（X,Y,Z,Rx,Ry,Rz）",
    variable=traj_type, value="TCP",
    command=_update_traj_labels_and_defaults
).pack_forget()

# 重新建立带 command 的两个单选按钮
for widget in list(type_frame.pack_slaves()):
    if isinstance(widget, tk.Radiobutton):
        widget.destroy()

tk.Radiobutton(
    type_frame, text="TCP（X,Y,Z,Rx,Ry,Rz）",
    variable=traj_type, value="TCP",
    command=_update_traj_labels_and_defaults
).pack(side=tk.LEFT, padx=8)

tk.Radiobutton(
    type_frame, text="关节（J1~J6）",
    variable=traj_type, value="JOINT",
    command=_update_traj_labels_and_defaults
).pack(side=tk.LEFT, padx=8)

btn_traj_input = tk.Frame(tab_traj)
btn_traj_input.pack(fill=tk.X, padx=10, pady=3)

tk.Button(
    btn_traj_input,
    text="检查并加入当前点",
    command=add_and_check_trajectory_point,
    width=22,
    bg="#2196F3",
    fg="white",
    font=("Microsoft YaHei", 10, "bold")
).pack(side=tk.LEFT, padx=3)

tk.Button(
    btn_traj_input,
    text="读取当前TCP并写入",
    command=read_current_tcp_to_traj,
    width=20
).pack(side=tk.LEFT, padx=3)

tk.Button(
    btn_traj_input,
    text="读取当前关节并写入",
    command=read_current_joints_to_traj,
    width=20
).pack(side=tk.LEFT, padx=3)

tk.Button(
    btn_traj_input,
    text="清空当前输入",
    command=clear_trajectory_input,
    width=16
).pack(side=tk.LEFT, padx=3)

tk.Label(
    tab_traj,
    text="输入一个点后：TCP 用 IK 判断可达；关节点不做检查，输入合法后直接加入。只有 TCP 检查通过的点或合法关节点才会加入下面列表。",
    fg="#555555"
).pack(anchor=tk.W, padx=15, pady=3)

frame_record = tk.LabelFrame(
    tab_traj,
    text="已检查通过的连续运动点（按加入顺序执行，可混合 TCP / 关节点）"
)
frame_record.pack(fill=tk.BOTH, expand=True, padx=10, pady=8)

record_text = tk.Text(frame_record, font=("Consolas", 10), height=10)
record_text.pack(fill=tk.BOTH, expand=True, padx=5, pady=5)

btn_record_frame = tk.Frame(tab_traj)
btn_record_frame.pack(fill=tk.X, padx=10, pady=4)

tk.Button(
    btn_record_frame, text="删除最后一点",
    command=delete_last_record, width=15
).pack(side=tk.LEFT, padx=3)

tk.Button(
    btn_record_frame, text="清空全部点",
    command=clear_records, width=15
).pack(side=tk.LEFT, padx=3)

tk.Button(
    btn_record_frame, text="导入轨迹",
    command=import_trajectory, width=14
).pack(side=tk.LEFT, padx=3)

tk.Button(
    btn_record_frame, text="执行整段连续运动",
    command=execute_recorded_trajectory,
    width=24,
    font=("Microsoft YaHei", 10, "bold"),
    bg="#4CAF50", fg="white"
).pack(side=tk.LEFT, padx=3)

tk.Label(
    tab_traj,
    text="执行：普通 TCP 首点 MoveJ、后续优先 MoveL；MoveL 失败直接用仿真已验证的 IK 解 MoveJ 兜底；末端特异点仅 J6 ±180°；关节点直接 MoveJ。实机不重复做轨迹预检。",
    fg="#555555"
).pack(anchor=tk.W, padx=15, pady=4)

# ---- 日志区 ----
frame_log = tk.LabelFrame(root, text="日志")
frame_log.pack(fill=tk.BOTH, expand=True, padx=10, pady=5)

text_log = scrolledtext.ScrolledText(frame_log, font=("Consolas", 10), height=8)
text_log.pack(fill=tk.BOTH, expand=True, padx=5, pady=5)

# ============================================================
# 启动
# ============================================================
log("机器人: " + robot.Name())
log("程序就绪。模式：RUNMODE_RUN_ROBOT + robot.Connect()")
log("单点：输入坐标 -> 检测可达性 -> 执行 MoveL/MoveJ")
log("目标关节：输入 J1~J6 -> 实机 MoveJ（不经过 TCP/Fanuc 转换和 IK）")
log("连续运动：支持导入仿真JSON；普通TCP使用仿真已验证IK（缺少时仅做单点SolveIK）；末端特异点跳过IK仅J6±180°；实机执行不重复轨迹预检；MoveL失败直接用仿真已验证IK解MoveJ兜底")

root.mainloop()

--- Python program 方向角计算 ---
import math
import tkinter as tk
from tkinter import ttk, messagebox

from robodk.robomath import Mat, Pose_2_Fanuc


# ============================================================
# 法兰坐标系 X+/Y+/Z+ -> RoboDK Fanuc/Motoman Rxyz
#
# 重要定义：
#   本程序现在不再只使用“末端朝向 Z 轴”计算姿态。
#   因为仅指定 Z+ 只能确定法兰朝向，不能确定绕 Z+ 的旋转。
#
#   现在可以同时输入：
#       X+ 在世界坐标中的方向
#       Y+ 在世界坐标中的方向
#       Z+ 在世界坐标中的方向
#
#   三个轴共同决定完整的法兰姿态。
#
#   如果只知道 Z+：
#       可以使用“Z+ + X+参考方向”模式，
#       程序会自动把 X+参考方向投影到垂直于 Z+ 的平面。
#
# 输出：
#   RoboDK Fanuc/Motoman [X,Y,Z,Rx,Ry,Rz]
#
# 单位：
#   输入向量：无单位，只表示方向
#   Rxyz：deg
# ============================================================


def vec_length(v):
    return math.sqrt(
        v[0] * v[0] +
        v[1] * v[1] +
        v[2] * v[2]
    )


def normalize(v):
    length = vec_length(v)

    if length < 1e-12:
        raise ValueError("方向向量不能为零向量")

    return (
        v[0] / length,
        v[1] / length,
        v[2] / length
    )


def dot(a, b):
    return (
        a[0] * b[0] +
        a[1] * b[1] +
        a[2] * b[2]
    )


def cross(a, b):
    return (
        a[1] * b[2] - a[2] * b[1],
        a[2] * b[0] - a[0] * b[2],
        a[0] * b[1] - a[1] * b[0]
    )


def scale(v, s):
    return (
        v[0] * s,
        v[1] * s,
        v[2] * s
    )


def sub(a, b):
    return (
        a[0] - b[0],
        a[1] - b[1],
        a[2] - b[2]
    )


def axis_to_rxyz(x_axis, y_axis, z_axis):
    """
    已知完整的法兰坐标系 X+/Y+/Z+ 在世界坐标中的方向，
    构造旋转矩阵并转换为 RoboDK Fanuc/Motoman Rxyz。
    """

    # 三个轴都归一化
    x_axis = normalize(x_axis)
    y_axis = normalize(y_axis)
    z_axis = normalize(z_axis)

    # 基本正交性检查
    xy = abs(dot(x_axis, y_axis))
    yz = abs(dot(y_axis, z_axis))
    zx = abs(dot(z_axis, x_axis))

    if max(xy, yz, zx) > 0.02:
        raise ValueError(
            "输入的 X+/Y+/Z+ 不是相互垂直的坐标轴。\n"
            "请检查三个方向向量。"
        )

    # 右手系检查：
    # X × Y 应该等于 Z
    cross_xy = normalize(cross(x_axis, y_axis))
    if dot(cross_xy, z_axis) < 0:
        raise ValueError(
            "输入的 X+/Y+/Z+ 不是右手坐标系。\n"
            "必须满足 X+ × Y+ = Z+。"
        )

    pose = Mat([
        [x_axis[0], y_axis[0], z_axis[0], 0],
        [x_axis[1], y_axis[1], z_axis[1], 0],
        [x_axis[2], y_axis[2], z_axis[2], 0],
        [0,         0,         0,         1]
    ])

    fanuc = Pose_2_Fanuc(pose)

    return (
        fanuc[3],
        fanuc[4],
        fanuc[5],
        pose
    )


def z_and_x_reference_to_rxyz(z_direction, x_reference):
    """
    已知 Z+ 方向，以及一个“X+参考方向”，
    自动构造完整右手坐标系。

    X+参考方向不要求本身严格垂直 Z+。
    程序会把它投影到垂直于 Z+ 的平面。
    """

    z_axis = normalize(z_direction)
    x_ref = normalize(x_reference)

    # X参考方向投影到垂直 Z+ 的平面
    x_axis = sub(
        x_ref,
        scale(z_axis, dot(x_ref, z_axis))
    )

    if vec_length(x_axis) < 1e-8:
        raise ValueError(
            "Z+ 与 X+参考方向平行或接近平行，"
            "无法确定滚转方向。"
        )

    x_axis = normalize(x_axis)

    # 右手系：X × Y = Z
    # 因此 Y = Z × X
    y_axis = normalize(cross(z_axis, x_axis))

    return axis_to_rxyz(x_axis, y_axis, z_axis)


def rotate_flange_z(pose, angle_deg):
    """绕法兰自身 Z+ 轴右手旋转；从 Z+ 端朝原点看，正角为逆时针。"""
    if not math.isfinite(angle_deg):
        raise ValueError("旋转角度必须是有限数字。")
    angle = math.radians(angle_deg)
    c, s = math.cos(angle), math.sin(angle)
    rotation = Mat([
        [c, -s, 0, 0],
        [s,  c, 0, 0],
        [0,  0, 1, 0],
        [0,  0, 0, 1]
    ])
    # 右乘表示绕局部轴旋转，而不是基座 Z 轴。
    rotated = pose * rotation
    values = Pose_2_Fanuc(rotated)
    return values[3], values[4], values[5], rotated


class DirectionToRxyzGUI:
    def __init__(self, root):
        self.root = root
        self.root.title("CR5 法兰坐标系 → RoboDK Rxyz")
        self.root.geometry("960x880")
        self.root.minsize(900, 800)

        self.mode = tk.StringVar(value="full")
        self.rotation_var = tk.StringVar(value="0")
        self.rotation_direction = tk.StringVar(value="顺时针")

        self.x_vars = [tk.StringVar() for _ in range(3)]
        self.y_vars = [tk.StringVar() for _ in range(3)]
        self.z_vars = [tk.StringVar() for _ in range(3)]

        self._build_ui()

        # 默认使用你目前讨论的方向。
        # 注意：这里给的是“法兰 Z+”，不是工具 Z-。
        self._set_axis(self.z_vars, 0, -1, 0)

        # 一组与 Z+=(0,-1,0) 配套的右手坐标系：
        # X+=(1,0,0)
        # Y+=(0,0,1)
        self._set_axis(self.x_vars, 1, 0, 0)
        self._set_axis(self.y_vars, 0, 0, 1)

        self.calculate()

    def _build_ui(self):
        ttk.Label(
            self.root,
            text="CR5 法兰坐标系 X+/Y+/Z+ → RoboDK Fanuc/Motoman Rxyz",
            font=("Microsoft YaHei UI", 16, "bold")
        ).pack(pady=(15, 5))

        ttk.Label(
            self.root,
            text=(
                "现在同时考虑红色 X+、绿色 Y+、蓝色 Z+。"
                "三根轴共同决定完整姿态。"
            ),
            font=("Microsoft YaHei UI", 10)
        ).pack(pady=(0, 12))

        # ====================================================
        # 模式选择
        # ====================================================
        mode_frame = ttk.LabelFrame(
            self.root,
            text="计算方式",
            padding=10
        )
        mode_frame.pack(fill="x", padx=18, pady=6)

        ttk.Radiobutton(
            mode_frame,
            text="完整坐标轴模式：输入 X+ / Y+ / Z+",
            variable=self.mode,
            value="full",
            command=self._update_mode
        ).pack(anchor="w")

        ttk.Radiobutton(
            mode_frame,
            text="方向 + 滚转参考模式：输入 Z+，再给一个 X+参考方向",
            variable=self.mode,
            value="zx",
            command=self._update_mode
        ).pack(anchor="w", pady=(5, 0))

        # ====================================================
        # 完整坐标轴输入
        # ====================================================
        self.full_frame = ttk.LabelFrame(
            self.root,
            text="1A. 法兰三个正方向（世界坐标）",
            padding=10
        )
        self.full_frame.pack(fill="x", padx=18, pady=6)

        self._build_axis_row(
            self.full_frame, "X+（红色）", self.x_vars, 0
        )
        self._build_axis_row(
            self.full_frame, "Y+（绿色）", self.y_vars, 1
        )
        self._build_axis_row(
            self.full_frame, "Z+（蓝色）", self.z_vars, 2
        )

        # ====================================================
        # Z+ + X参考输入
        # ====================================================
        self.zx_frame = ttk.LabelFrame(
            self.root,
            text="1B. Z+方向 + X+滚转参考",
            padding=10
        )

        self._build_axis_row(
            self.zx_frame, "Z+（蓝色）", self.z_vars, 0
        )
        self._build_axis_row(
            self.zx_frame, "X+参考（红色）", self.x_vars, 1
        )

        # ====================================================
        # 快速测试
        # ====================================================
        preset_frame = ttk.LabelFrame(
            self.root,
            text="快速测试",
            padding=10
        )
        preset_frame.pack(fill="x", padx=18, pady=6)

        ttk.Button(
            preset_frame,
            text="图中方向：Z+=(0,-1,0)",
            command=self.preset_current
        ).pack(side="left", padx=5)

        ttk.Button(
            preset_frame,
            text="Z+=+X",
            command=lambda: self.preset_z(1, 0, 0)
        ).pack(side="left", padx=5)

        ttk.Button(
            preset_frame,
            text="Z+=+Y",
            command=lambda: self.preset_z(0, 1, 0)
        ).pack(side="left", padx=5)

        ttk.Button(
            preset_frame,
            text="Z+=+Z",
            command=lambda: self.preset_z(0, 0, 1)
        ).pack(side="left", padx=5)

        rotation_frame = ttk.LabelFrame(
            self.root, text="末端追加旋转（绕法兰自身 Z 轴）", padding=10
        )
        rotation_frame.pack(fill="x", padx=18, pady=6)
        ttk.Label(rotation_frame, text="角度（度，非负）：").grid(row=0, column=0)
        ttk.Entry(rotation_frame, textvariable=self.rotation_var, width=12).grid(
            row=0, column=1, padx=8
        )
        ttk.Combobox(
            rotation_frame, textvariable=self.rotation_direction,
            values=("顺时针", "逆时针"), state="readonly", width=10
        ).grid(row=0, column=2, padx=8)
        ttk.Label(
            rotation_frame,
            text="观察方向：从法兰 Z+ 端朝原点看。每次均相对输入姿态计算，不累加。"
        ).grid(row=1, column=0, columnspan=3, sticky="w", pady=(8, 0))

        # ====================================================
        # 操作
        # ====================================================
        button_frame = ttk.Frame(self.root)
        button_frame.pack(pady=10)

        ttk.Button(
            button_frame,
            text="计算 Rxyz",
            command=self.calculate
        ).pack(side="left", padx=8)

        ttk.Button(
            button_frame,
            text="清空",
            command=self.clear
        ).pack(side="left", padx=8)

        # ====================================================
        # 结果
        # ====================================================
        result_frame = ttk.LabelFrame(
            self.root,
            text="2. 计算结果",
            padding=10
        )
        result_frame.pack(
            fill="both",
            expand=True,
            padx=18,
            pady=6
        )

        self.result_text = tk.Text(
            result_frame,
            font=("Consolas", 11),
            wrap="none"
        )
        self.result_text.pack(
            side="left",
            fill="both",
            expand=True
        )

        scrollbar = ttk.Scrollbar(
            result_frame,
            orient="vertical",
            command=self.result_text.yview
        )
        scrollbar.pack(side="right", fill="y")

        self.result_text.configure(
            yscrollcommand=scrollbar.set
        )

        ttk.Label(
            self.root,
            text=(
                "注意：仅一个 Z+ 方向不能唯一确定 Rxyz；"
                "必须再规定 X+/Y+ 的滚转方向。"
            ),
            font=("Microsoft YaHei UI", 9)
        ).pack(pady=(3, 12))

    def _build_axis_row(self, parent, title, vars_, row):
        ttk.Label(
            parent,
            text=title,
            width=18,
            font=("Microsoft YaHei UI", 10, "bold")
        ).grid(
            row=row,
            column=0,
            padx=(4, 10),
            pady=5,
            sticky="w"
        )

        for i, (axis_name, var) in enumerate(
            zip(["X", "Y", "Z"], vars_)
        ):
            ttk.Label(
                parent,
                text=axis_name
            ).grid(
                row=row,
                column=1 + i * 2,
                padx=(3, 4)
            )

            ttk.Entry(
                parent,
                textvariable=var,
                width=12,
                justify="center"
            ).grid(
                row=row,
                column=2 + i * 2,
                padx=(0, 12)
            )

    def _update_mode(self):
        if self.mode.get() == "full":
            self.zx_frame.pack_forget()
            self.full_frame.pack(
                fill="x",
                padx=18,
                pady=6,
                before=self._find_widget("快速测试")
            )
        else:
            self.full_frame.pack_forget()
            self.zx_frame.pack(
                fill="x",
                padx=18,
                pady=6,
                before=self._find_widget("快速测试")
            )

    def _find_widget(self, text):
        # 简单返回当前界面中的第一个 LabelFrame，
        # 这里只用于控制布局；找不到时返回 self
        for widget in self.root.winfo_children():
            if isinstance(widget, ttk.LabelFrame):
                if widget.cget("text") == text:
                    return widget
        return self.root

    def _set_axis(self, vars_, x, y, z):
        vars_[0].set(str(x))
        vars_[1].set(str(y))
        vars_[2].set(str(z))

    def preset_current(self):
        self._set_axis(self.z_vars, 0, -1, 0)
        self._set_axis(self.x_vars, 1, 0, 0)
        self._set_axis(self.y_vars, 0, 0, 1)
        self.mode.set("full")
        self._update_mode()
        self.calculate()

    def preset_z(self, x, y, z):
        self._set_axis(self.z_vars, x, y, z)

        # 根据 Z+ 自动寻找一个简单的 X+参考方向
        if abs(x) < 0.9:
            self._set_axis(self.x_vars, 1, 0, 0)
        else:
            self._set_axis(self.x_vars, 0, 1, 0)

        self.mode.set("zx")
        self._update_mode()
        self.calculate()

    def _read_vec(self, vars_, name):
        try:
            values = [
                float(var.get().strip())
                for var in vars_
            ]
        except (ValueError, AttributeError):
            raise ValueError(
                "%s 的三个分量必须全部是数字。" % name
            )

        if not all(math.isfinite(v) for v in values):
            raise ValueError(
                "%s 不能包含 NaN 或无穷值。" % name
            )

        return tuple(values)

    def calculate(self):
        try:
            if self.mode.get() == "full":
                x_axis = self._read_vec(self.x_vars, "X+")
                y_axis = self._read_vec(self.y_vars, "Y+")
                z_axis = self._read_vec(self.z_vars, "Z+")
                rx, ry, rz, pose = axis_to_rxyz(x_axis, y_axis, z_axis)
                mode_text = "完整坐标轴模式：直接使用输入的 X+/Y+/Z+"
            else:
                z_axis = self._read_vec(self.z_vars, "Z+")
                x_ref = self._read_vec(self.x_vars, "X+参考")
                rx, ry, rz, pose = z_and_x_reference_to_rxyz(z_axis, x_ref)
                x_axis = (pose[0,0], pose[1,0], pose[2,0])
                y_axis = (pose[0,1], pose[1,1], pose[2,1])
                z_axis = (pose[0,2], pose[1,2], pose[2,2])
                mode_text = "Z+ + X+参考模式：X+参考已投影到垂直 Z+ 的平面"

            # 处理旋转角度
            angle_deg = float(self.rotation_var.get().strip())
            if not math.isfinite(angle_deg) or angle_deg < 0:
                raise ValueError("旋转角度必须是非负有限数字。")
            signed_angle = -angle_deg if self.rotation_direction.get() == "顺时针" else angle_deg
            rx, ry, rz, pose = rotate_flange_z(pose, signed_angle)

            # 提取旋转后的轴向量
            x_axis = (pose[0,0], pose[1,0], pose[2,0])
            y_axis = (pose[0,1], pose[1,1], pose[2,1])
            z_axis = (pose[0,2], pose[1,2], pose[2,2])

            # ===== 新增：回填姿态到输入框，实现连续累加 =====
            self._set_axis(self.x_vars, x_axis[0], x_axis[1], x_axis[2])
            self._set_axis(self.y_vars, y_axis[0], y_axis[1], y_axis[2])
            self._set_axis(self.z_vars, z_axis[0], z_axis[1], z_axis[2])
            # 切换模式到“完整坐标轴模式”，以便显示三个轴
            self.mode.set("full")
            self._update_mode()
            # ===================================================

            mode_text += (
                "\n追加旋转：%s %.6f°（从 Z+ 端朝原点看）"
                "\n绕法兰局部 Z 轴，右手角度 = %+.6f°"
                % (self.rotation_direction.get(), angle_deg, signed_angle)
            )

            result = (
                "========================================\n"
                "CR5 法兰坐标系 → RoboDK Rxyz\n"
                "========================================\n\n"
                "【计算模式】\n"
                "%s\n\n"
                "【最终法兰坐标轴（世界坐标）】\n"
                "X+ = (%+.6f, %+.6f, %+.6f)\n"
                "Y+ = (%+.6f, %+.6f, %+.6f)\n"
                "Z+ = (%+.6f, %+.6f, %+.6f)\n\n"
                "【旋转矩阵 R】\n"
                "[ %+.6f  %+.6f  %+.6f ]\n"
                "[ %+.6f  %+.6f  %+.6f ]\n"
                "[ %+.6f  %+.6f  %+.6f ]\n\n"
                "【RoboDK Fanuc/Motoman】\n"
                "Rx = %+.6f deg\n"
                "Ry = %+.6f deg\n"
                "Rz = %+.6f deg\n\n"
                "【可直接用于 RoboDK 的位姿】\n"
                "[0, 0, 0, %.6f, %.6f, %.6f]\n\n"
                "【轴方向说明】\n"
                "红色箭头 = X+\n"
                "绿色箭头 = Y+\n"
                "蓝色箭头 = Z+\n\n"
                "注意：\n"
                "这里的 Z+ 就是你图片中确认的法兰蓝色箭头。\n"
                "因此不再对输入 Z+ 取反。\n"
                % (
                    mode_text,
                    x_axis[0], x_axis[1], x_axis[2],
                    y_axis[0], y_axis[1], y_axis[2],
                    z_axis[0], z_axis[1], z_axis[2],
                    pose[0,0], pose[0,1], pose[0,2],
                    pose[1,0], pose[1,1], pose[1,2],
                    pose[2,0], pose[2,1], pose[2,2],
                    rx, ry, rz,
                    rx, ry, rz
                )
            )

            self.result_text.delete("1.0", tk.END)
            self.result_text.insert("1.0", result)

        except Exception as e:
            messagebox.showerror("计算失败", "%s: %s" % (type(e).__name__, e))

    def clear(self):
        self.rotation_var.set("0")
        self.rotation_direction.set("顺时针")
        for var in (
            self.x_vars +
            self.y_vars +
            self.z_vars
        ):
            var.set("")

        self.result_text.delete("1.0", tk.END)


def main():
    root = tk.Tk()

    DirectionToRxyzGUI(root)

    root.mainloop()


if __name__ == "__main__":
    main()

--- Python program test ---
#!/usr/bin/env python3
# -*- coding: utf-8 -*-
"""原点 -> P1 -> P2 -> P3 -> P4(奇异点) -> P5 -> P6 -> P7 -> P8(奇异点) -> P9 -> P10
单步运动测试（GUI，TCP 坐标版；带【台面/地面】碰撞预检 + 自动换解）

P1 / P2 = **轨迹3（连续轨迹3.json）的第 1、2 个点**，原样就是 TCP（法兰 Fanuc 六数）；
P3 / P5 / P6 / P7 / P9 / P10 = 后续新增的普通 TCP 点；**P4 / P8 = 奇异点**（只走关节运动）：
    P1  =  500.0,   0.0, 300.0, 180.0,  0.0,   0.0
    P2  =    0.0, -775.0, 300.0, -90.0, 0.0, 180.0
    P3  =  100.0, -775.0, 300.0, -90.0, 0.0, 180.0
    P4  =  100.0, -775.0, 300.0, -90.0, 0.0,   0.0   ← ★ 奇异点：不做 IK，只让 J6 转 ±180°
    P5  =    0.0, -775.0, 300.0,  90.0, 0.0,   0.0
    P6  =    0.0, -770.0, 300.0, 180.0, 0.0,   0.0
    P7  =  100.0, -770.0, 300.0, 180.0, 0.0,   0.0
    P8  =  100.0, -770.0, 300.0, 180.0, 0.0, 180.0   ← ★ 奇异点：不做 IK，只让 J6 转 ±180°
    P9  =    0.0, -770.0, 300.0, 180.0, 0.0, 180.0
    P10 = -500.0,    0.0, 300.0, 180.0, 0.0,   0.0
起点 = 原点（关节 0,0,0,0,0,0；按习惯机械臂开跑前就在原点）。

【★ P4 特殊处理（照抄 机械臂法兰真实运动.py 的“末端特异点/直接控制关节运动”选项）】
    该点的位姿在腕部奇异处，TCP 逆解会退化 ⇒ **不做 TCP 运动、不做 SolveIK**：
      · 取【当前实际关节】原样，只把 J6 加上 P4_J6_DELTA（默认 +180°）
      · 角度规范化到 (-180, 180]（照抄参考脚本第 512-514 行）
      · 仍然做一次碰撞预检（关节目标 ⇒ 无解可换，只测这一条）
      · 然后直接 MoveJ(关节目标) —— 即“直接控制关节运动”

【十段运动 & 延时】① 原点->P1  ② P1->P2  ③ P2->P3  ④ P3->P4(仅 J6 ±180°)  ⑤ P4->P5
                    ⑥ P5->P6   ⑦ P6->P7  ⑧ P7->P8(仅 J6 ±180°)  ⑨ P8->P9  ⑩ P9->P10 ；
                    ★ 每段运动之前额外延时 SEG_DELAY=2 秒。

【★ 碰撞预检（照抄 机械臂TCP仿真.py）】
    障碍物只取两个：
        安装台_650x650x80mm   —— 台面
        地面_禁止穿越          —— 地面
    ✗ 不管磨砂圆盘      ✗ 不考虑末端工具（参考脚本里“工具 × 障碍物”那段按要求省略）

    ★★ 关键：不拒绝任务，而是【换解】——
       robot.SolveIK_All(target) 枚举全部逆解
         ⇒ 每个解归一化到 ±180°，J6 再试 0 / −1 / +1 圈，滤掉超关节限位的
         ⇒ 按 _obstacle_posture_key 排序（肘部相对台面越高越优先）
         ⇒ 逐个 robot.MoveJ_Test(起点, 候选, minstep=1°)（碰撞检查已开）
         ⇒ 取【第一个通过】的候选作为本段的执行目标 ✓✓
       ⇒ 于是"预检通过的构型" 就是 "实际执行的构型"，且能绕开台面/地面继续运动。

【单步逻辑】严格照抄 机械臂法兰真实运动.py 的 execute_joint_target：
    ensure_connected() -> RDK.setRunMode(RUNMODE_RUN_ROBOT) -> robot.setSpeed(...) -> robot.MoveJ(target)
    ✗ 不开 30004   ✗ 不用 robot.Joints()/Busy()/setPoseFrame/setPoseTool
★ StoppedError 兜底仍保留（驱动会假报 'Robot not connected'，本环境常态）。

★ 运行前提：机械臂在原点；路径清空；手放急停上；RoboDK 已打开并加载【含台子和地面】的工作站。
"""
from robodk.robolink import *
from robodk.robomath import *
import tkinter as tk
from tkinter import scrolledtext
import math
import queue
import threading
import time

ROBOT_SPEED = 20.0       # ★ 速度：2026-09-28 按要求恢复到 20.0（此前减半为 10.0）
SEG_DELAY = 0.5          # ★ 每段运动前的延时（秒）：2026-09-28 按要求 2.0 → 0.5
NL = chr(10)

# ---- ★ 碰撞预检（只查台面 + 地面）----
COLLISION_OBSTACLES = ('安装台_650x650x80mm', '地面_禁止穿越')
TABLE_NAME = '安装台_650x650x80mm'
CHECK_MINSTEP_DEG = 1.0   # 与参考脚本的主检测粒度一致
CHECK_ENABLED = True      # 默认开启；GUI 可切换
MAX_CANDIDATES_TRY = 24   # 最多试多少个候选解（防御性上限）

# ---- 起点（关节；机械臂开跑前就在原点）----
ORIGIN_JOINTS = [0.0, 0.0, 0.0, 0.0, 0.0, 0.0]

# ---- 两个目标点：轨迹3 的第 1、2 点，TCP（法兰 Fanuc）原样照抄 ----
P1_TCP = [500.0, 0.0, 300.0, 180.0, 0.0, 0.0]
P2_TCP = [0.0, -775.0, 300.0, -90.0, 0.0, 180.0]
P3_TCP = [100.0, -775.0, 300.0, -90.0, 0.0, 180.0]   # ★ 新增第 3 点（本次要求）
# ★★ 第 4 点 = 【奇异点】：不要走 TCP 运动（其 IK 在腕部奇异处会退化）
#    照抄 机械臂法兰真实运动.py 的"末端特异点"处理：完全跳过 SolveIK，
#    保持 J1~J5 不变，执行时只让 J6 转 ±180°（默认 +180°）。
P4_TCP = [100.0, -775.0, 300.0, -90.0, 0.0, 0.0]     # 仅作记录/日志，不用于 IK
P4_IS_SINGULAR = True
P4_J6_DELTA = 180.0                                  # ±180（+180 = 参考脚本默认）
# ★ 第 5 点：普通 TCP 点（回到正常 TCP 运动 + 碰撞预检换解）
P5_TCP = [0.0, -775.0, 300.0, 90.0, 0.0, 0.0]
# ★ 第 6 点：普通 TCP 点
P6_TCP = [0.0, -770.0, 300.0, 180.0, 0.0, 0.0]
# ★ 第 7 点：普通 TCP 点
P7_TCP = [100.0, -770.0, 300.0, 180.0, 0.0, 0.0]
# ★★ 第 8 点 = 【奇异点】（与第 4 点同类）：只差 Rz 0→180 ⇒ 直接控制关节，仅让 J6 转 ±180°
P8_TCP = [100.0, -770.0, 300.0, 180.0, 0.0, 180.0]   # 仅作记录/日志，不用于 IK
P8_IS_SINGULAR = True
P8_J6_DELTA = 180.0                                  # ±180（+180 = 参考脚本默认）
# ★ 第 9 / 10 点：普通 TCP 点
P9_TCP = [0.0, -770.0, 300.0, 180.0, 0.0, 180.0]
P10_TCP = [-500.0, 0.0, 300.0, 180.0, 0.0, 0.0]

# ---- 碰撞预检结果缓存（生命周期 = 单次预检；每次 _enable_obstacle_checks 清空）----
_plan_cache = {}

RDK = None
robot = None
text_log = None
run_btn = None
status_var = None
check_var = None
_running = False
_connected = False
_msg_q = queue.Queue()


def log(s):
    print(s, flush=True)
    _msg_q.put(str(s))


def _pump():
    try:
        while True:
            s = _msg_q.get_nowait()
            if text_log is not None:
                text_log.insert(tk.END, s + NL)
                text_log.see(tk.END)
    except queue.Empty:
        pass
    root.after(80, _pump)


# ============================================================
# 连接（照抄法兰脚本 ensure_connected）
# ============================================================
def init_robot():
    global RDK, robot
    if RDK is None:
        RDK = Robolink()
    if robot is None:
        robot = RDK.Item('', ITEM_TYPE_ROBOT)
    return robot is not None and robot.Valid()


def ensure_connected():
    global _connected
    if _connected:
        return True
    if not init_robot():
        log("!! 未在 RoboDK 站点里找到机器人（ITEM_TYPE_ROBOT）")
        return False
    try:
        robot.Connect()
        time.sleep(1.5)
        status, msg = robot.ConnectedState()
        log("连接状态: %s, %s" % (status, msg))
        if status != ROBOTCOM_READY:
            log("机器人未就绪：status=%s msg=%s" % (status, msg))
            _connected = False
            return False
        RDK.setRunMode(RUNMODE_RUN_ROBOT)
        log("RunMode: %s" % RDK.RunMode())
        _connected = True
        return True
    except Exception as e:  # noqa: BLE001
        log("连接失败: %s: %s" % (type(e).__name__, e))
        return False


# ============================================================
# 坐标换算（照抄法兰脚本的数学，一字不改）
# ============================================================
def _tool_mat():
    try:
        t = robot.PoseTool()
        return t if t is not None else eye(4)
    except Exception:
        return eye(4)


def fanuc_to_pose(x, y, z, rx, ry, rz):
    """【法兰】位姿(Fanuc) -> 当前工具下的 TCP 位姿（参考坐标系中）。"""
    return Fanuc_2_Pose([x, y, z, rx, ry, rz]) * _tool_mat()


def _sim_joints():
    q = list(robot.SimulatorJoints())
    return [float(v) for v in q[:6]] if len(q) >= 6 else None


def _fmt(vals):
    return ('X=%+.3f Y=%+.3f Z=%+.3f Rx=%+.3f Ry=%+.3f Rz=%+.3f'
            % (vals[0], vals[1], vals[2], vals[3], vals[4], vals[5]))


def _fmtq(q):
    return ("J1=%+.4f J2=%+.4f J3=%+.4f J4=%+.4f J5=%+.4f J6=%+.4f" % tuple(list(q)[:6]))


def read_current():
    if not ensure_connected():
        return
    try:
        q = _sim_joints()
        log("当前位置（SimulatorJoints）：" + (_fmtq(q) if q else '(读不到 6 个值)'))
    except Exception as e:  # noqa: BLE001
        log("读取失败: %s: %s" % (type(e).__name__, e))


# ============================================================
# ★ 碰撞预检（台面 + 地面）—— 照抄 机械臂TCP仿真.py 的换解逻辑
# ============================================================
def _cache_key_joints(q):
    return tuple(round(float(v), 3) for v in q[:6])


def _movej_test_cached(start, end, minstep_deg):
    """robot.MoveJ_Test 的缓存包装（照抄参考脚本）。"""
    key = ('movej_test', _cache_key_joints(start), _cache_key_joints(end),
           round(float(minstep_deg), 6))
    if key not in _plan_cache:
        _plan_cache[key] = robot.MoveJ_Test(start, end, minstep_deg=minstep_deg)
    elif _plan_cache[key] == 0:
        robot.setJoints(list(end[:6]))
    return _plan_cache[key]


def _collision_details():
    pairs = RDK.CollisionPairs()
    return '；'.join('%s[连杆%d] 与 %s[连杆%d]' % (a.Name(), ia, b.Name(), ib)
                     for a, b, ia, ib in pairs) or '路径碰撞或关节不可行'


def _enable_obstacle_checks():
    """照抄参考脚本，但按要求【不给末端工具配碰撞对】。
       必须在 RUNMODE_SIMULATE 下调用。"""
    if RDK.RunMode() != RUNMODE_SIMULATE:
        raise RuntimeError('障碍物碰撞预检仅允许在仿真模式执行。')
    _plan_cache.clear()
    for name in COLLISION_OBSTACLES:
        obstacle = RDK.Item(name, ITEM_TYPE_OBJECT)
        if not obstacle.Valid():
            raise RuntimeError('缺少障碍物模型：%s，请加载包含台子和地面的工作站。' % name)
        if name == TABLE_NAME:
            # 固定底座与台面本来就接触，不参与判定（照抄参考脚本）
            if RDK.setCollisionActivePair(COLLISION_OFF, robot, obstacle, 0, 0) != 1:
                raise RuntimeError('无法配置安装台与固定底座的接触关系。')
        for link in range(1, 7):
            if RDK.setCollisionActivePair(COLLISION_ON, robot, obstacle, link, 0) != 1:
                raise RuntimeError('无法启用 %s 与连杆%d 的碰撞检查。' % (name, link))
        # ★ 参考脚本这里还有 “for tool in RDK.ItemList(ITEM_TYPE_TOOL)”
        #   —— 本次按要求【不考虑末端工具】，故省略。
    RDK.setCollisionActive(COLLISION_ON)


def _obstacle_posture_key(q, reference=None):
    """照抄参考脚本：优先"肘部（连杆3）离台面更高"的构型；再优先离当前关节更近的。"""
    height = 0.0
    try:
        table = RDK.Item(TABLE_NAME, ITEM_TYPE_OBJECT)
        if table.Valid():
            elbow = invH(table.PoseAbs()) * robot.PoseAbs() * robot.JointPoses(q)[3]
            height = float(elbow.Pos()[2])
    except Exception:
        height = 0.0
    ref = reference or [0.0] * 6
    return (-round(height, 6), sum((v - r) ** 2 for v, r in zip(q, ref)), tuple(q))


def _tcp_target_to_flange(pose):
    """TCP 位姿 -> 法兰位姿（照抄参考脚本 机械臂TCP仿真.py 第 758-760 行）。
    ★ 必须做这一步：SolveIK / SolveIK_All 要的是【法兰】位姿，而 fanuc_to_pose
      返回的是【TCP】位姿（已乘过工具矩阵）。漏掉这一步会解不出逆解。"""
    return robot.PoseFrame() * pose * invH(robot.PoseTool())


def _singular_j6_target(start_joints, delta):
    """构造"末端特异点"的关节目标：保持 J1~J5 不变，只让 J6 转 ±delta。

    照抄参考脚本 机械臂法兰真实运动.py 的“末端特异点/直接控制关节运动”做法：
      · 完全跳过 SolveIK（该位姿在腕部奇异处，逆解会退化）
      · J6 加 ±delta（默认 ±180°）
      · 角度规范化到 (-180, 180]（参考脚本第 512-514 行）
    """
    q = [float(v) for v in start_joints[:6]]
    q[5] += delta
    q = [((v + 180.0) % 360.0) - 180.0 for v in q]
    return [180.0 if v <= -180.0 else v for v in q]


def _run_singular_segment(tag, p_label, delta, tcp_for_log, seg_index, seg_total, fallback_start=None):
    """执行一个"末端特异点"段：跳过 IK，仅 J6 ±delta，仍然做碰撞预检。

    返回 (是否放行, 起点关节, 目标关节)。
    """
    log("")
    log("--- 段 %d / %d：%s（奇异点：跳过 IK，仅 J6 %+g°）---" % (seg_index, seg_total, tag, delta))
    log("    %s  目标（仅记录）%s" % (p_label, _fmt(tcp_for_log)))
    log("    ★ 该点标记为末端特异点 ⇒ 不做 TCP 逆解；保持 J1~J5 不变，只让 J6 转 %+g°" % delta)
    log("      （做法照抄 机械臂法兰真实运动.py 的“末端特异点/直接控制关节运动”选项）")
    log("延时 %.1f 秒 ..." % SEG_DELAY)
    time.sleep(SEG_DELAY)

    start = _sim_joints() or fallback_start or list(ORIGIN_JOINTS)
    target = _singular_j6_target(start, delta)
    log("      起点关节：%s" % _fmtq(start))
    log("      目标关节：%s   （J6 %+.4f° → %+.4f°）" % (_fmtq(target), start[5], target[5]))

    allow, chosen = _do_segment_check(start, target, "段%d %s（仅 J6 %+g°）" % (seg_index, tag, delta))
    return allow, start, (chosen if chosen else target)


def _ik_candidates(pose, reference):
    """枚举目标位姿的全部可用关节解（照抄参考脚本 _trajectory_start_candidates）。"""
    try:
        solutions = robot.SolveIK_All(_tcp_target_to_flange(pose))   # ★ 法兰位姿
    except Exception as e:  # noqa: BLE001
        log("      SolveIK_All 异常：%s: %s" % (type(e).__name__, e))
        return []
    try:
        lower, upper, _ = robot.JointLimits()
        lower = [float(v) for v in list(lower)[:6]]
        upper = [float(v) for v in list(upper)[:6]]
    except Exception:
        lower = [-360.0] * 6
        upper = [360.0] * 6

    candidates = []
    for solution in solutions:
        q = [((float(v) + 180.0) % 360.0) - 180.0 for v in list(solution)[:6]]
        if len(q) != 6:
            continue
        for turns6 in (0, -1, 1):
            cand = q[:]
            cand[5] += 360.0 * turns6
            if all(lower[j] <= cand[j] <= upper[j] for j in range(6)):
                if not any(max(abs(a - b) for a, b in zip(cand, old)) < 1e-6 for old in candidates):
                    candidates.append(cand)
    # 同一姿态保留"接近当前圈数"的表示（照抄参考脚本）
    for q in candidates[:]:
        try:
            nearest = [min((v + 360 * k for k in range(
                int(math.ceil((lower[j] - v) / 360.0)),
                int(math.floor((upper[j] - v) / 360.0)) + 1)),
                key=lambda a: abs(a - reference[j]))
                for j, v in enumerate(q)]
        except Exception:
            continue
        if not any(max(abs(a - b) for a, b in zip(nearest, old)) < 1e-6 for old in candidates):
            candidates.append(nearest)
    return sorted(candidates, key=lambda q: _obstacle_posture_key(q, reference))


def _check_segment(start_joints, target, tag):
    """在【仿真模式】下为 start_joints -> target 这一段【挑一个不撞台面/地面的构型】。

    target 可以是关节列表（6 个数，此时无解可换）或位姿（Mat，此时枚举全部逆解换解）。
    返回 (ok, chosen_joints, message)。
    ★ 无论成败都把 RunMode 恢复原值；只动模型，不发真机指令。
    """
    saved_mode = RDK.RunMode()
    saved_joints = None
    try:
        RDK.setRunMode(RUNMODE_SIMULATE)
        _enable_obstacle_checks()
        try:
            saved_joints = [float(v) for v in robot.Joints()][:6]
        except Exception:
            saved_joints = None

        # ---- 目标是关节（如"回原点"）：没有候选可换，只测这一条 ----
        if isinstance(target, (list, tuple)) and len(target) == 6:
            robot.setJoints(list(start_joints[:6]))
            status = _movej_test_cached(start_joints, list(target), CHECK_MINSTEP_DEG)
            if status == 0:
                return True, list(target), '通过（关节目标，status=0）'
            return False, None, '不通过（status=%s）：%s' % (status, _collision_details())

        # ---- 目标是位姿：枚举全部逆解，按肘高排序，逐个测 ----
        cands = _ik_candidates(target, start_joints)
        log("      逆解候选 %d 个（SolveIK_All，已转法兰位姿），按【肘部离台面高度】排序后逐个做 MoveJ_Test …" % len(cands))
        if not cands:
            # ★ 兜底：让 RoboDK 自己解（MoveJ_Test 也接受位姿）——TCP 位姿 / 法兰位姿各试一次
            log("      枚举为空 ⇒ 兜底：直接让 RoboDK 自己解（MoveJ_Test 接受位姿）")
            for label, tgt in (('TCP 位姿', target), ('法兰位姿', _tcp_target_to_flange(target))):
                try:
                    robot.setJoints(list(start_joints[:6]))
                    st = robot.MoveJ_Test(start_joints, tgt, minstep_deg=CHECK_MINSTEP_DEG)
                except Exception as e:  # noqa: BLE001
                    log("      %s 兜底异常：%s: %s" % (label, type(e).__name__, e))
                    continue
                if st == 0:
                    try:
                        end = [float(v) for v in robot.Joints()][:6]
                    except Exception:
                        end = None
                    log("      ✓ %s 兜底通过（status=0），终点关节 %s"
                        % (label, _fmtq(end) if end else '(读不到)'))
                    return True, end, '通过（%s 兜底，RoboDK 自解，status=0）' % label
                log("      ✗ %s 兜底未通过 status=%s" % (label, st))
            return False, None, '没有可用逆解（SolveIK_All 无解，且两种位姿兜底都未通过）'

        tried = 0
        for cand in cands[:MAX_CANDIDATES_TRY]:
            tried += 1
            try:
                robot.setJoints(list(start_joints[:6]))
            except Exception:
                pass
            status = _movej_test_cached(start_joints, cand, CHECK_MINSTEP_DEG)
            h = _obstacle_posture_key(cand, start_joints)[0]
            if status == 0:
                log("      ✓ 第 %d 个候选通过（肘部相对台面 %.1f mm）：%s" % (tried, -h, _fmtq(cand)))
                return True, cand, '通过（第 %d/%d 个候选，status=0）' % (tried, len(cands))
            log("      ✗ 第 %d 个候选未通过 status=%s（肘部 %.1f mm）" % (tried, status, -h))
        return False, None, '全部 %d 个候选都未通过：%s' % (tried, _collision_details())
    except Exception as e:  # noqa: BLE001
        return False, None, '预检异常：%s: %s' % (type(e).__name__, e)
    finally:
        try:
            if saved_joints is not None:
                robot.setJoints(saved_joints)     # 只影响模型
        except Exception:
            pass
        try:
            RDK.setRunMode(saved_mode)            # ★ 必须切回原模式
        except Exception:
            pass


# ============================================================
# 单步运动（照抄 execute_joint_target，并保留你自己的 StoppedError 兜底）
# ============================================================
def _stationary(a, b, tol=0.05):
    return bool(a) and bool(b) and max(abs(x - y) for x, y in zip(a, b)) <= tol


def _move_one(target, tag, target_joints=None):
    """单步 MoveJ。

    照抄 execute_joint_target 的四步；但**保留** 机械臂TCP真实运动.py 第 618-632 行的兜底：
    驱动会假报 `StoppedError: Robot not connected`（指令其实已发出，报错发生在"等待完成"阶段），
    此环境里是常态，不能当失败。
    判据改用【RoboDK 模型关节 SimulatorJoints】（连接真机时模型与真机同步）
    —— 不读 30004、不碰任何端口，因此不会再被端口占用拖死。
      ① 若给了 target_joints（原点那种）：模型到位即算完成；
      ② 否则要求"确实动过 + 已停稳"：证明指令执行过且这一段落停住了。
    """
    q_before = _sim_joints()
    log("  发送 MoveJ -> %s" % tag)
    RDK.setRunMode(RUNMODE_RUN_ROBOT)
    robot.setSpeed(ROBOT_SPEED)
    try:
        robot.MoveJ(target)                      # ← 照抄：不加兜底、不读反馈
        log("  ✓ %s：MoveJ 命令已发送并返回" % tag)
        return True
    except StoppedError as exc:
        if str(exc).strip() != 'Robot not connected':
            raise                                # 其它 StoppedError 一律照抄原样上抛
    log("  ⚠ 驱动返回 'Robot not connected'（已知假报警；发生在等待完成阶段）")
    log("     判定中：用模型关节（SimulatorJoints）确认这一段是否真的走完 …")
    for attempt in range(10):
        time.sleep(0.3)
        a = _sim_joints()
        time.sleep(0.3)
        b = _sim_joints()
        if not _stationary(a, b):
            continue                             # 还在动，继续等
        if target_joints is not None:
            if max(abs(x - y) for x, y in zip(b, target_joints)) <= 0.5:
                log("  ✓ %s：模型关节已到目标且停稳 %s ⇒ 计为完成，不重发" % (tag, _fmtq(b)))
                return True
        elif q_before is not None and max(abs(x - y) for x, y in zip(b, q_before)) > 0.05:
            log("  ✓ %s：已停稳且确实动过（%s → %s）⇒ 计为完成，不重发"
                % (tag, _fmtq(q_before), _fmtq(b)))
            return True
    raise RuntimeError("驱动报 'Robot not connected'，但模型关节既未到位也未显示『动过且停稳』"
                       "（第 %d 次尝试后）⇒ 判定为真失败" % (10 + 1))


def _do_segment_check(start_joints, target, tag):
    """执行一段前的碰撞预检（含换解）；返回 (是否放行, 本段要执行的关节目标)。"""
    if not CHECK_ENABLED:
        log("  （碰撞预检已关闭，跳过）")
        return True, (list(target) if isinstance(target, (list, tuple)) and len(target) == 6 else None)
    log("  碰撞预检（台面 + 地面，含换解）：%s" % tag)
    ok, chosen, msg = _check_segment(start_joints, target, tag)
    if ok:
        log("  ✓ %s：预检通过 —— %s" % (tag, msg))
        return True, chosen
    log("  ✗ %s：预检未通过 ⇒ 本段不执行，以避免碰撞" % tag)
    log("     原因：%s" % msg)
    return False, None


def _worker():
    global _running
    try:
        log("")
        log("=" * 64)
        log("单步测试（TCP 坐标版 + 台面/地面碰撞预检/换解）：原点 -> 轨迹3 P1 -> 轨迹3 P2")
        log("速度 %.1f ｜ 每段运动前延时 %.1f 秒 ｜ 碰撞预检 %s"
            % (ROBOT_SPEED, SEG_DELAY, "开" if CHECK_ENABLED else "关"))
        log("障碍物：%s（不含磨砂圆盘；不含末端工具）" % ', '.join(COLLISION_OBSTACLES))
        log("=" * 64)
        if not ensure_connected():
            raise RuntimeError("连接未建立，取消")

        try:
            q0 = _sim_joints()
            if q0:
                log("起始位置（SimulatorJoints）：" + _fmtq(q0))
                log("距离原点最大偏差 = %.4f°" % max(abs(v) for v in q0))
        except Exception as e:  # noqa: BLE001
            log("读取起始位置失败（不阻断）：%s: %s" % (type(e).__name__, e))

        origin = list(ORIGIN_JOINTS)   # ★ 原点是【关节】目标（不是位姿！）
        p1 = fanuc_to_pose(*P1_TCP)
        p2 = fanuc_to_pose(*P2_TCP)
        p3 = fanuc_to_pose(*P3_TCP)
        p5 = fanuc_to_pose(*P5_TCP)
        p6 = fanuc_to_pose(*P6_TCP)
        p7 = fanuc_to_pose(*P7_TCP)
        p9 = fanuc_to_pose(*P9_TCP)
        p10 = fanuc_to_pose(*P10_TCP)

        # ---- 段 1 / 10：当前位置 -> 原点 -> P1 ----
        log("")
        log("--- 段 1 / 10：原点 -> P1 ---")
        log("    原点目标（关节）%s" % _fmtq(ORIGIN_JOINTS))
        log("    P1  目标 %s" % _fmt(P1_TCP))
        log("延时 %.1f 秒 ..." % SEG_DELAY)
        time.sleep(SEG_DELAY)

        # ★ 碰撞预检：回到原点这一段（关节目标，无解可换）
        seg_start = _sim_joints() or list(ORIGIN_JOINTS)
        allow0, chosen0 = _do_segment_check(seg_start, origin, "段1a 当前 -> 原点")
        if not allow0:
            log("")
            log("!! 回到原点这一段预检未通过 ⇒ 取消（未发送任何运动指令）")
            raise RuntimeError("段1a（回原点）碰撞预检未通过")
        _move_one(origin, "原点", ORIGIN_JOINTS)

        # ★ 碰撞预检：原点 -> P1（位姿目标 ⇒ 会枚举逆解并换解）
        seg_start = _sim_joints() or list(ORIGIN_JOINTS)
        allow1, chosen1 = _do_segment_check(seg_start, p1, "段1b 原点 -> P1")
        if not allow1:
            log("")
            log("!! 段1 因碰撞预检未通过而取消（未发送任何运动指令）")
            raise RuntimeError("段1 碰撞预检未通过")
        # ★ 执行【预检选中的那个构型】，保证"检查过的解 = 走的解"
        _move_one(chosen1 if chosen1 else p1, "P1（轨迹3 第1点）", chosen1)

        # ---- 段 2 / 10：P1 -> P2 ----
        log("")
        log("--- 段 2 / 10：P1 -> P2 ---")
        log("    P2  目标 %s" % _fmt(P2_TCP))
        log("延时 %.1f 秒 ..." % SEG_DELAY)
        time.sleep(SEG_DELAY)

        seg_start2 = _sim_joints() or chosen1 or list(ORIGIN_JOINTS)
        allow2, chosen2 = _do_segment_check(seg_start2, p2, "段2 P1 -> P2")
        if not allow2:
            log("")
            log("!! 段2 因碰撞预检未通过而取消（未发送任何运动指令）")
            raise RuntimeError("段2 碰撞预检未通过")
        _move_one(chosen2 if chosen2 else p2, "P2（轨迹3 第2点）", chosen2)

        # ---- 段 3 / 10：P2 -> P3 ----
        log("")
        log("--- 段 3 / 10：P2 -> P3 ---")
        log("    P3  目标 %s" % _fmt(P3_TCP))
        log("延时 %.1f 秒 ..." % SEG_DELAY)
        time.sleep(SEG_DELAY)

        seg_start3 = _sim_joints() or chosen2 or list(ORIGIN_JOINTS)
        allow3, chosen3 = _do_segment_check(seg_start3, p3, "段3 P2 -> P3")
        if not allow3:
            log("")
            log("!! 段3 因碰撞预检未通过而取消（未发送任何运动指令）")
            raise RuntimeError("段3 碰撞预检未通过")
        _move_one(chosen3 if chosen3 else p3, "P3（第3点）", chosen3)

        # ---- 段 4 / 10：P3 -> P4（★ 奇异点：不走 TCP 运动，直接控制关节 —— 只让 J6 转 ±180°）----
        allow4, seg_start4, j6_target = _run_singular_segment(
            "P3 -> P4", "P4", P4_J6_DELTA, P4_TCP, 4, 8, fallback_start=chosen3)
        if not allow4:
            log("")
            log("!! 段4 因碰撞预检未通过而取消（未发送任何运动指令）")
            raise RuntimeError("段4 碰撞预检未通过")
        _move_one(j6_target, "P4（第4点，仅 J6 %+g°）" % P4_J6_DELTA, j6_target)

        # ---- 段 5 / 10：P4 -> P5（普通 TCP 点 ⇒ 回到 TCP 运动 + 碰撞预检换解）----
        log("")
        log("--- 段 5 / 10：P4 -> P5 ---")
        log("    P5  目标 %s" % _fmt(P5_TCP))
        log("延时 %.1f 秒 ..." % SEG_DELAY)
        time.sleep(SEG_DELAY)

        seg_start5 = _sim_joints() or chosen4 or j6_target or list(ORIGIN_JOINTS)
        allow5, chosen5 = _do_segment_check(seg_start5, p5, "段5 P4 -> P5")
        if not allow5:
            log("")
            log("!! 段5 因碰撞预检未通过而取消（未发送任何运动指令）")
            raise RuntimeError("段5 碰撞预检未通过")
        _move_one(chosen5 if chosen5 else p5, "P5（第5点）", chosen5)

        # ---- 段 6 / 10：P5 -> P6（普通 TCP 点）----
        log("")
        log("--- 段 6 / 10：P5 -> P6 ---")
        log("    P6  目标 %s" % _fmt(P6_TCP))
        log("延时 %.1f 秒 ..." % SEG_DELAY)
        time.sleep(SEG_DELAY)

        seg_start6 = _sim_joints() or chosen5 or list(ORIGIN_JOINTS)
        allow6, chosen6 = _do_segment_check(seg_start6, p6, "段6 P5 -> P6")
        if not allow6:
            log("")
            log("!! 段6 因碰撞预检未通过而取消（未发送任何运动指令）")
            raise RuntimeError("段6 碰撞预检未通过")
        _move_one(chosen6 if chosen6 else p6, "P6（第6点）", chosen6)

        # ---- 段 7 / 10：P6 -> P7（普通 TCP 点）----
        log("")
        log("--- 段 7 / 10：P6 -> P7 ---")
        log("    P7  目标 %s" % _fmt(P7_TCP))
        log("延时 %.1f 秒 ..." % SEG_DELAY)
        time.sleep(SEG_DELAY)

        seg_start7 = _sim_joints() or chosen6 or list(ORIGIN_JOINTS)
        allow7, chosen7 = _do_segment_check(seg_start7, p7, "段7 P6 -> P7")
        if not allow7:
            log("")
            log("!! 段7 因碰撞预检未通过而取消（未发送任何运动指令）")
            raise RuntimeError("段7 碰撞预检未通过")
        _move_one(chosen7 if chosen7 else p7, "P7（第7点）", chosen7)

        # ---- 段 8 / 10：P7 -> P8（★ 奇异点：不走 TCP 运动，直接控制关节 —— 只让 J6 转 ±180°）----
        allow8, seg_start8, j6_target8 = _run_singular_segment(
            "P7 -> P8", "P8", P8_J6_DELTA, P8_TCP, 8, 8, fallback_start=chosen7)
        if not allow8:
            log("")
            log("!! 段8 因碰撞预检未通过而取消（未发送任何运动指令）")
            raise RuntimeError("段8 碰撞预检未通过")
        _move_one(j6_target8, "P8（第8点，仅 J6 %+g°）" % P8_J6_DELTA, j6_target8)

        # ---- 段 9 / 10：P8 -> P9（普通 TCP 点）----
        log("")
        log("--- 段 9 / 10：P8 -> P9 ---")
        log("    P9  目标 %s" % _fmt(P9_TCP))
        log("延时 %.1f 秒 ..." % SEG_DELAY)
        time.sleep(SEG_DELAY)

        seg_start9 = _sim_joints() or j6_target8 or list(ORIGIN_JOINTS)
        allow9, chosen9 = _do_segment_check(seg_start9, p9, "段9 P8 -> P9")
        if not allow9:
            log("")
            log("!! 段9 因碰撞预检未通过而取消（未发送任何运动指令）")
            raise RuntimeError("段9 碰撞预检未通过")
        _move_one(chosen9 if chosen9 else p9, "P9（第9点）", chosen9)

        # ---- 段 10 / 10：P9 -> P10（普通 TCP 点）----
        log("")
        log("--- 段 10 / 10：P9 -> P10 ---")
        log("    P10 目标 %s" % _fmt(P10_TCP))
        log("延时 %.1f 秒 ..." % SEG_DELAY)
        time.sleep(SEG_DELAY)

        seg_start10 = _sim_joints() or chosen9 or list(ORIGIN_JOINTS)
        allow10, chosen10 = _do_segment_check(seg_start10, p10, "段10 P9 -> P10")
        if not allow10:
            log("")
            log("!! 段10 因碰撞预检未通过而取消（未发送任何运动指令）")
            raise RuntimeError("段10 碰撞预检未通过")
        _move_one(chosen10 if chosen10 else p10, "P10（第10点）", chosen10)

        log("")
        log("=" * 64)
        try:
            q = _sim_joints()
            if q:
                log("结束位置（SimulatorJoints）：" + _fmtq(q))
        except Exception:
            pass
        log("全部完成 ✓")
        log("=" * 64)
    except Exception as e:  # noqa: BLE001
        import traceback
        log("")
        log("!! 中断：%s: %s" % (type(e).__name__, e))
        for line in traceback.format_exc().rstrip().splitlines():
            log("   " + line)
        log("（照抄原脚本行为：不自动重发运动；请检查机械臂与报警）")
    finally:
        _running = False
        try:
            RDK.setRunMode(RUNMODE_RUN_ROBOT)     # 收尾确保回到真机模式
        except Exception:
            pass
        try:
            run_btn.configure(state=tk.NORMAL, text="启动运动")
            status_var.set("就绪")
        except Exception:
            pass


def start_motion():
    global _running, CHECK_ENABLED
    if _running:
        log("已在运行中，忽略本次点击")
        return
    try:
        CHECK_ENABLED = bool(check_var.get())
    except Exception:
        pass
    _running = True
    run_btn.configure(state=tk.DISABLED, text="运行中 ...")
    status_var.set("运行中")
    log("")
    log("########## 启动运动 ##########")
    threading.Thread(target=_worker, daemon=True).start()


# ============================================================
# GUI
# ============================================================
root = tk.Tk()
root.title("RoboDK - 原点→P1→P2→P3→P4(奇异点)→P5→P6→P7→P8(奇异点)→P9→P10 单步测试")
root.geometry("1060x740")
root.resizable(True, True)

frame_top = tk.LabelFrame(root, text="测试内容（单步 / TCP 坐标 / 台面+地面碰撞预检，含自动换解）")
frame_top.pack(fill=tk.X, padx=10, pady=6)
tk.Label(frame_top, anchor=tk.W, justify=tk.LEFT,
         text=("段1:原点->P1  段2:P1->P2  段3:P2->P3  段4:P3->P4(仅J6±180°)  段5:P4->P5  段6:P5->P6  段7:P6->P7  段8:P7->P8(仅J6±180°)  段9:P8->P9  段10:P9->P10" + NL
               + "        每段运动前延时 " + str(SEG_DELAY) + " 秒" + NL
               + "P1（轨迹3 第1点）= 500.0, 0.0, 300.0, 180.0, 0.0, 0.0              （TCP / 法兰 Fanuc）" + NL
               + "P2（轨迹3 第2点）= 0.0, -775.0, 300.0, -90.0, 0.0, 180.0" + NL
               + "P3（第3点）      = 100.0, -775.0, 300.0, -90.0, 0.0, 180.0" + NL
               + "P4（★奇异点）    = 100.0, -775.0, 300.0, -90.0, 0.0, 0.0   ← 不做 TCP 逆解" + NL
               + "P5（第5点）      = 0.0, -775.0, 300.0, 90.0, 0.0, 0.0      ← 普通 TCP 点" + NL
               + "P6（第6点）      = 0.0, -770.0, 300.0, 180.0, 0.0, 0.0     ← 普通 TCP 点" + NL
               + "P7（第7点）      = 100.0, -770.0, 300.0, 180.0, 0.0, 0.0   ← 普通 TCP 点" + NL
               + "P8（★奇异点）    = 100.0, -770.0, 300.0, 180.0, 0.0, 180.0 ← 不做 TCP 逆解" + NL
               + "P9（第9点）      = 0.0, -770.0, 300.0, 180.0, 0.0, 180.0   ← 普通 TCP 点" + NL
               + "P10（第10点）    = -500.0, 0.0, 300.0, 180.0, 0.0, 0.0     ← 普通 TCP 点" + NL
               + "   ★ P4 / P8 走“直接控制关节运动”：保持 J1~J5 不变，只让 J6 转 " + str(P4_J6_DELTA)
               + "°，然后直接 MoveJ(关节)" + NL
               + "★ 碰撞预检：障碍物 = 安装台_650x650x80mm（台面）+ 地面_禁止穿越（地面）" + NL
               + "   做法照抄 机械臂TCP仿真.py：SolveIK_All 枚举全部逆解 → 按“肘部离台面高度”排序" + NL
               + "   → 逐个 MoveJ_Test（1° 粒度、碰撞开）→ 取第一个通过的构型去执行 ✓"),
         font=("Microsoft YaHei", 10)).pack(fill=tk.X, padx=8, pady=4)

frame_btn = tk.LabelFrame(root, text="操作")
frame_btn.pack(fill=tk.X, padx=10, pady=6)
run_btn = tk.Button(frame_btn, text="启动运动", width=18, bg="#4CAF50", fg="white",
                    font=("Microsoft YaHei", 11, "bold"), command=start_motion)
run_btn.pack(side=tk.LEFT, padx=8, pady=8)
check_var = tk.BooleanVar(value=True)
tk.Checkbutton(frame_btn, text="碰撞预检（台面+地面，含换解）", variable=check_var,
               font=("Microsoft YaHei", 10)).pack(side=tk.LEFT, padx=6, pady=8)
tk.Button(frame_btn, text="读取当前位置", width=16, font=("Microsoft YaHei", 10),
          command=lambda: threading.Thread(target=read_current, daemon=True).start()
          ).pack(side=tk.LEFT, padx=6, pady=8)
tk.Button(frame_btn, text="清空日志", width=12, font=("Microsoft YaHei", 10),
          command=lambda: text_log.delete("1.0", tk.END)).pack(side=tk.LEFT, padx=6, pady=8)
status_var = tk.StringVar(value="就绪")
tk.Label(frame_btn, textvariable=status_var, anchor=tk.W, fg="#555",
         font=("Microsoft YaHei", 10)).pack(side=tk.LEFT, padx=16)

frame_log = tk.LabelFrame(root, text="日志")
frame_log.pack(fill=tk.BOTH, expand=True, padx=10, pady=6)
text_log = scrolledtext.ScrolledText(frame_log, font=("Consolas", 10), height=20)
text_log.pack(fill=tk.BOTH, expand=True, padx=5, pady=5)

log("程序就绪。模式：RUNMODE_RUN_ROBOT + robot.Connect()；碰撞预检在 RUNMODE_SIMULATE 下进行")
log("测试 = 单步：原点 -> P1 -> P2 -> P3 -> P4(奇异点) -> P5 -> P6 -> P7 -> P8(奇异点) -> P9 -> P10（TCP 坐标）")
log("P1 = 500.0, 0.0, 300.0, 180.0, 0.0, 0.0")
log("P2 = 0.0, -775.0, 300.0, -90.0, 0.0, 180.0")
log("P3 = 100.0, -775.0, 300.0, -90.0, 0.0, 180.0")
log("P4 = 100.0, -775.0, 300.0, -90.0, 0.0, 0.0   ★奇异点：不做 IK，保持 J1~J5，只让 J6 转 %+g°" % P4_J6_DELTA)
log("P5 = 0.0, -775.0, 300.0, 90.0, 0.0, 0.0      （普通 TCP 点）")
log("P6 = 0.0, -770.0, 300.0, 180.0, 0.0, 0.0     （普通 TCP 点）")
log("P7 = 100.0, -770.0, 300.0, 180.0, 0.0, 0.0   （普通 TCP 点）")
log("P8 = 100.0, -770.0, 300.0, 180.0, 0.0, 180.0  ★奇异点：不做 IK，保持 J1~J5，只让 J6 转 %+g°" % P8_J6_DELTA)
log("P9 = 0.0, -770.0, 300.0, 180.0, 0.0, 180.0   （普通 TCP 点）")
log("P10 = -500.0, 0.0, 300.0, 180.0, 0.0, 0.0    （普通 TCP 点）")
log("★ 碰撞预检障碍物：安装台_650x650x80mm（台面）、地面_禁止穿越（地面）；不含磨砂圆盘、不含末端工具")
log("★ 预检不通过时会自动换解（SolveIK_All 全部逆解 → 肘高排序 → 逐个 MoveJ_Test）")
log("★ 运行前请确认：机械臂在原点、路径清空、手放急停上、工作站里已加载台子和地面")
log("")
_pump()
root.mainloop()

--- Python program 机械臂法兰真实运动_改名修复前_20261014_114144_改名修复前_20261014_114144 ---
# -*- coding: utf-8 -*-
"""
RoboDK 实机运动控制 —— 【法兰坐标版】（不把末端工具算进去）
- 单点：法兰位姿(Fanuc 格式) 输入 -> IK 检测 -> MoveL/MoveJ 执行
- 连续轨迹：法兰位姿/关节点列表 -> 逐点 IK 检测 -> MoveJ+MoveL 序列
- 关节点直通：J1~J6 -> 实机 MoveJ（不经 TCP/IK，本来就是法兰无关）

坐标约定（与 机械臂TCP真实运动.py 的唯一区别）：
  本脚本输入/显示/记录的都是【法兰】(flange) 位姿 —— 不含末端工具。
  RoboDK 的 SolveIK / MoveL / MoveJ 一律按 TCP 解释位姿，所以：
    * 运动前：TCP目标 = 法兰 × 当前工具(PoseTool)   [fanuc_to_pose 里做]
    * 读取时：法兰   = invH(PoseFrame) × SolveFK(Joints)   [完全不含工具]
  ⇒ 换工具不需要改本脚本的任何坐标；工具只在最后一次换算里出现，且会在日志里打印。

⚠️ 与 TCP 版的数据不通用：TCP版导出的 JSON 里存的是 TCP 坐标，直接导入本脚本
   会整体偏移一个工具量。请只用本脚本自己导出的 JSON。

模式：RUNMODE_RUN_ROBOT + robot.Connect()
"""

from robodk.robolink import *
from robodk.robomath import *
import tkinter as tk
from tkinter import ttk, scrolledtext, filedialog
import time
import math
import json
import itertools

ROBOT_SPEED = 10.0       # ★ 速度：已按 2026-09-27 要求从 20.0 减半（原值 20.0）
NL = chr(10)

# ============================================================
# 连续运动逻辑的常量与预检缓存（整段移植自仿真脚本，算法未改动）
# ============================================================
ALLOW_MOTION = True
MOVEJ_FALLBACK_MAX_DEVIATION_MM = 500.0  # MoveL失败后，MoveJ轨迹允许偏离TCP直线段的最大距离

# ============================================================
# 碰撞判断排除清单（本阶段：磨砂圆盘暂不参与碰撞判断）
# ============================================================
# 工位对象名只要【包含】下面任一关键字，就显式关掉它与机器人和所有工具的
# 碰撞判断（只关这一个对象的配对，安装台/地面等其它障碍物不受影响）。
# 当前命中的工位对象：磨砂圆柱_R180_H40（即磨砂圆盘）。
# 要恢复它的碰撞判断：把这里改成空元组 EXCLUDED_COLLISION_KEYWORDS = () 即可。
# 注意：RoboDK 默认就会对工位内对象做碰撞判断，所以这里是"显式关掉"，
# 而不是"不再添加"。
EXCLUDED_COLLISION_KEYWORDS = ('磨砂',)

# ============================================================
# 预检结果缓存（性能优化：分支重试不重复计算，判定结果不变）
# ============================================================
# 缓存生命周期 = 单次预检规划：_enable_obstacle_checks() 在每次进入预检时
# 清空缓存，因此障碍物/工作站状态的任何变化都会在下一次预检中即时生效。
_plan_cache = {}

def _cache_key_joints(q):
    return tuple(round(float(v), 3) for v in q[:6])

def _cache_key_pose(pose):
    return tuple(tuple(round(float(v), 6) for v in row) for row in pose.rows)

def _movej_test_cached(start, end, minstep_deg):
    """robot.MoveJ_Test 的缓存包装，返回值与直接调用完全一致。
    成功时与原调用一样把仿真关节停在终点；失败路径的规划器只依赖局部
    关节变量（不读取此时的模型关节状态），无需复现失败的副作用。"""
    key = ('movej_test', _cache_key_joints(start), _cache_key_joints(end),
           round(float(minstep_deg), 6))
    if key not in _plan_cache:
        _plan_cache[key] = robot.MoveJ_Test(start, end, minstep_deg=minstep_deg)
    elif _plan_cache[key] == 0:
        robot.setJoints(list(end[:6]))
    return _plan_cache[key]

RDK = Robolink()

def _tool_mat():
    """当前工具位姿（TCP 相对法兰）。取不到就退回单位阵（等价于以法兰为 TCP）。"""
    try:
        t = robot.PoseTool()
        return t if t is not None else eye(4)
    except Exception:
        return eye(4)

def fanuc_to_pose(x, y, z, rx, ry, rz):
    """【法兰】位姿(Fanuc) -> 当前工具下的 TCP 位姿。

    操作员给的是法兰坐标；RoboDK 的 SolveIK/MoveL/MoveJ 都要 TCP，
    所以在入口处做一次 法兰 × 工具，之后所有既有代码原样复用。
    """
    flange = Fanuc_2_Pose([x, y, z, rx, ry, rz])
    return flange * _tool_mat()

def pose_to_fanuc(pose):
    return Pose_2_Fanuc(pose)

def _joints6():
    """读取当前关节（6 个）。

    ⚠️ 本环境**不能用 robot.Joints()**：实机模式下它会去读真机驱动，超时后 RoboDK
    只返回 1×1 的 [[0]]（屏幕上是 "Robot connection failed timed out: Working..."），
    后面任何按 6 个用的地方都会 IndexError。已验证的实机脚本（机械臂TCP真实运动.py）
    一律用 SimulatorJoints()（RoboDK 模型姿态；连接真机时模型与真机同步）。
    读不到 6 个就明确报错，不再让 IndexError 冒到上层。
    """
    try:
        q = list(robot.SimulatorJoints())
    except Exception as exc:
        raise RuntimeError(f'读取当前关节失败：{type(exc).__name__}: {exc}')
    if len(q) < 6:
        raise RuntimeError(f'读取当前关节失败：SimulatorJoints 只返回 {len(q)} 个值 {q}；'
                           '请确认 RoboDK 里机器人已连接、模型姿态显示正常。')
    return [float(v) for v in q[:6]]


def current_flange_pose():
    """当前【法兰】位姿（当前参考坐标系下，不含工具）。

    等价于 invH(PoseFrame) × Pose，但不引入工具量，因此工具的改动不会影响读数。
    """
    return invH(robot.PoseFrame()) * robot.SolveFK(_joints6())

# ---- 名称适配：仿真脚本的连续运动逻辑使用下面两个名字 ----
# 这是零改动的转发（法兰边界仍然只在 _tool_mat / fanuc_to_pose / pose_to_fanuc /
# current_flange_pose 里实现，坐标数学一律没有改动）。
def fanuc_values_to_pose(x, y, z, rx, ry, rz):
    """等同 fanuc_to_pose：法兰位姿(Fanuc) -> 当前工具下的 TCP 位姿。"""
    return fanuc_to_pose(x, y, z, rx, ry, rz)

def pose_to_fanuc_values(pose):
    """等同 pose_to_fanuc：位姿 -> Fanuc 六数。"""
    return pose_to_fanuc(pose)

# ---- 获取机器人 ----
robot = RDK.Item('', ITEM_TYPE_ROBOT)
if not robot.Valid():
    raise Exception("未找到机器人")

# ---- 全局变量 ----
text_points = None
text_log = None
record_text = None
entries_single = None
entries_joint = None
move_type = None
trajectory_records = []
_connected = False
simulation_running = False   # 连续运动是否正在运行（移植自仿真脚本）

# ============================================================
# 日志
# ============================================================
def log(s):
    """写三处：stdout + 单点日志(text_log) + 连续运动日志(traj_log_output/traj_status_var)。"""
    print(s)
    if text_log:
        try:
            text_log.insert(tk.END, str(s) + NL)
            text_log.see(tk.END)
        except Exception:
            pass
    try:
        traj_log_output.insert(tk.END, str(s) + NL)
        traj_log_output.see(tk.END)
    except Exception:
        pass
    try:
        if str(s).strip():
            traj_status_var.set(str(s))
    except Exception:
        pass
    try:
        root.update_idletasks()
    except Exception:
        pass

# ============================================================
# 连接（只连一次，复用）
# ============================================================
def ensure_connected():
    global _connected
    if _connected:
        return True
    try:
        robot.Connect()
        time.sleep(1.5)
        status, msg = robot.ConnectedState()
        log("连接状态: %s, %s" % (status, msg))
        RDK.setRunMode(RUNMODE_RUN_ROBOT)
        log("RunMode: %s" % RDK.RunMode())
        if status < 0:
            _connected = False
            log("机器人连接未建立，状态=%s：%s" % (status, msg))
            return False
        _connected = True
        return True
    except Exception as e:
        log("连接失败: %s" % e)
        return False

# ============================================================
# 解析坐标
# ============================================================
def parse_points():
    if not text_points:
        return []
    raw = text_points.get("1.0", tk.END)
    points = []
    for line in raw.strip().split(NL):
        line = line.strip()
        if not line or line.startswith("#"):
            continue
        try:
            vals = [float(v.strip()) for v in line.split(",")]
            if len(vals) >= 6:
                points.append(vals[:6])
        except ValueError:
            pass
    return points

# ============================================================
# 读取当前位置
# ============================================================
def read_current(entries=None):
    try:
        pose = current_flange_pose()
        v = pose_to_fanuc(pose)
        log("")
        log("当前法兰（不含工具）：X=%.3f Y=%.3f Z=%.3f Rx=%.3f Ry=%.3f Rz=%.3f" % tuple(v[:6]))
    except Exception as e:
        log("读取失败：%s" % e)

def fill_current(entries=None):
    try:
        pose = current_flange_pose()
        v = pose_to_fanuc(pose)
        if entries:
            for e, val in zip(entries, v):
                e.delete(0, tk.END)
                e.insert(0, "%.3f" % val)
        log("当前法兰（不含工具）已填入")
    except Exception as e:
        log("读取失败：%s" % e)

# ============================================================
# IK 检测
# 注意：SolveIK 显式使用当前 Tool + Reference，和 MoveL/MoveJ 保持一致。
# ============================================================
def check_ik_single(entries=None):
    if not entries:
        return
    try:
        values = [float(e.get()) for e in entries]
    except ValueError:
        log("输入无效")
        return

    x, y, z, rx, ry, rz = values
    target = fanuc_to_pose(x, y, z, rx, ry, rz)
    log("")
    log("目标：X=%.3f Y=%.3f Z=%.3f Rx=%.3f Ry=%.3f Rz=%.3f" % (x, y, z, rx, ry, rz))

    try:
        tool_pose = robot.PoseTool()
        frame_pose = robot.PoseFrame()
        joints = robot.SolveIK(target, tool=tool_pose, reference=frame_pose)
        if joints is None:
            log("IK 不可达")
        else:
            q = joints.list()
            if len(q) < 6:
                log("IK 返回关节数量异常：%d，原始数据=%r" % (len(q), q))
                return
            log("IK 可达")
            log("  关节：J1=%.2f J2=%.2f J3=%.2f J4=%.2f J5=%.2f J6=%.2f" % tuple(q[:6]))
    except Exception as e:
        log("检测失败：%s" % e)

def check_all_ik():
    points = parse_points()
    if not points:
        log("没有有效点")
        return

    log("")
    log("========== 检测全部 %d 个点 ==========" % len(points))
    all_ok = True
    for i, p in enumerate(points):
        try:
            target = fanuc_to_pose(*p)
            joints = robot.SolveIK(target, tool=robot.PoseTool(), reference=robot.PoseFrame())
            if joints is None:
                log("  P%d: 不可达" % (i+1))
                all_ok = False
            else:
                q = joints.list()
                if len(q) < 6:
                    raise ValueError("IK 返回关节数量异常: %d, raw=%r" % (len(q), q))
                log("  P%d: 可达  J1=%.1f J2=%.1f J3=%.1f J4=%.1f J5=%.1f J6=%.1f" % (i+1, *q[:6]))
        except Exception as e:
            log("  P%d: 检测失败 %s" % (i+1, e))
            all_ok = False
    if all_ok:
        log("全部 %d 个点可达" % len(points))
    else:
        log("存在不可达点，执行时会跳过")

# ============================================================
# 执行单点
# ============================================================
def execute_single(entries=None, mtype="MoveL"):
    if not entries:
        return
    try:
        values = [float(e.get()) for e in entries]
    except ValueError:
        log("输入无效")
        return

    x, y, z, rx, ry, rz = values
    target = fanuc_to_pose(x, y, z, rx, ry, rz)
    log("")
    log("目标：X=%.3f Y=%.3f Z=%.3f Rx=%.3f Ry=%.3f Rz=%.3f" % (x, y, z, rx, ry, rz))

    try:
        tool_pose = robot.PoseTool()
        frame_pose = robot.PoseFrame()
        joints = robot.SolveIK(target, tool=tool_pose, reference=frame_pose)
        if joints is None:
            log("IK 不可达，取消执行")
            return
        q = joints.list()
        if len(q) < 6:
            log("IK 返回关节数量异常：%d，取消执行；原始数据=%r" % (len(q), q))
            return
        log("IK 可达：J1=%.2f J2=%.2f J3=%.2f J4=%.2f J5=%.2f J6=%.2f" % tuple(q[:6]))
    except Exception as e:
        log("IK 检查失败：%s" % e)
        return

    if not ensure_connected():
        return

